(* IEC 61131-3 sources: 2026_Projet_YGO_ExcavatriceDragage/TOOLS/TEST_AUTO_CI/RESULTS/L_SIMULATION/tests (part 6) *)

(* ---- test_sim_operator_joystick.st ---- *)
(* T418 integration : vrais SimBench, FB_Joystick et homing, aucune logique machine remplacee.
   Temps explicite par scan : le DSL STruCpp interdit ADVANCE_TIME dans FOR. *)
SETUP
VAR
    bench : FB_SimBench;
    joy : FB_Joystick;
    home : FB_CycleMachineHoming;
    cfg : ST_fbJoystick_Cfg;
    diagOk : ST_Diag_Device;
    nx : INT := 5000;
    ny : INT := 5000;
    raw1 : UDINT;
    raw2 : UDINT;
    sourceSelected : BOOL;
    selectedX : INT;
    selectedY : INT;
    selectedButton : BOOL;
    previousButton : BOOL;
    buttonEdges : INT;
END_VAR
END_SETUP
TEST 'TC-T418-INT-001 Geste complet avec vrai joystick'
nx := 5000; ny := 5000; raw1 := 0; raw2 := 0; previousButton := FALSE; buttonEdges := 0;
bench.Enable := TRUE; joy.Enable := TRUE; joy.ArmingPermit := TRUE; diagOk.Operational := TRUE;
joy.BusCanOpenOP := diagOk; joy.JoystickOP := diagOk; home.Enable := TRUE; home.BootReady := TRUE;
home.Mode := E_Mode.MAINT_N1; home.BucketOffsetValid := TRUE; home.WinchesMechanicallyStopped := TRUE;
ADVANCE_TIME(10000000);
bench(RawPosM1 := raw1, RawPosM2 := raw2);
joy(RawX := bench.Operator.JoyXRaw_ANA1, RawY := bench.Operator.JoyYRaw_ANA2, RawButton := bench.Operator.JoyBtnRaw, Cfg := cfg, NeutralXMem := nx, NeutralYMem := ny);
home(DeadmanArmed := joy.DeadmanArmed, JoystickDeflected := NOT joy.AtNeutralXY, JoystickPull := joy.AxisCmdY.DirectionPositive, JoystickPush := joy.AxisCmdY.DirectionNegative, BtnValidation := bench.Operator.JoyBtnRaw);
IF bench.Operator.JoyBtnRaw AND NOT previousButton THEN buttonEdges := buttonEdges + 1; END_IF; previousButton := bench.Operator.JoyBtnRaw;
bench.SimJoystickRight_Fwd_MAINT_Active := TRUE;
ADVANCE_TIME(10000000);
bench(RawPosM1 := raw1, RawPosM2 := raw2);
joy(RawX := bench.Operator.JoyXRaw_ANA1, RawY := bench.Operator.JoyYRaw_ANA2, RawButton := bench.Operator.JoyBtnRaw, Cfg := cfg, NeutralXMem := nx, NeutralYMem := ny);
home(DeadmanArmed := joy.DeadmanArmed, JoystickDeflected := NOT joy.AtNeutralXY, JoystickPull := joy.AxisCmdY.DirectionPositive, JoystickPush := joy.AxisCmdY.DirectionNegative, BtnValidation := bench.Operator.JoyBtnRaw);
IF bench.Operator.JoyBtnRaw AND NOT previousButton THEN buttonEdges := buttonEdges + 1; END_IF; previousButton := bench.Operator.JoyBtnRaw;
ASSERT_EQ(bench.Operator.JoyXRaw_ANA1, 5000, 'Neutre pendant pre-appui');
ADVANCE_TIME(10000000);
bench(RawPosM1 := raw1, RawPosM2 := raw2);
joy(RawX := bench.Operator.JoyXRaw_ANA1, RawY := bench.Operator.JoyYRaw_ANA2, RawButton := bench.Operator.JoyBtnRaw, Cfg := cfg, NeutralXMem := nx, NeutralYMem := ny);
home(DeadmanArmed := joy.DeadmanArmed, JoystickDeflected := NOT joy.AtNeutralXY, JoystickPull := joy.AxisCmdY.DirectionPositive, JoystickPush := joy.AxisCmdY.DirectionNegative, BtnValidation := bench.Operator.JoyBtnRaw);
IF bench.Operator.JoyBtnRaw AND NOT previousButton THEN buttonEdges := buttonEdges + 1; END_IF; previousButton := bench.Operator.JoyBtnRaw;
ASSERT_EQ(bench.Operator.JoyXRaw_ANA1, 5000, 'Neutre pendant pre-appui');
ADVANCE_TIME(10000000);
bench(RawPosM1 := raw1, RawPosM2 := raw2);
joy(RawX := bench.Operator.JoyXRaw_ANA1, RawY := bench.Operator.JoyYRaw_ANA2, RawButton := bench.Operator.JoyBtnRaw, Cfg := cfg, NeutralXMem := nx, NeutralYMem := ny);
home(DeadmanArmed := joy.DeadmanArmed, JoystickDeflected := NOT joy.AtNeutralXY, JoystickPull := joy.AxisCmdY.DirectionPositive, JoystickPush := joy.AxisCmdY.DirectionNegative, BtnValidation := bench.Operator.JoyBtnRaw);
IF bench.Operator.JoyBtnRaw AND NOT previousButton THEN buttonEdges := buttonEdges + 1; END_IF; previousButton := bench.Operator.JoyBtnRaw;
ASSERT_EQ(bench.Operator.JoyXRaw_ANA1, 5000, 'Neutre pendant pre-appui');
ADVANCE_TIME(10000000);
bench(RawPosM1 := raw1, RawPosM2 := raw2);
joy(RawX := bench.Operator.JoyXRaw_ANA1, RawY := bench.Operator.JoyYRaw_ANA2, RawButton := bench.Operator.JoyBtnRaw, Cfg := cfg, NeutralXMem := nx, NeutralYMem := ny);
home(DeadmanArmed := joy.DeadmanArmed, JoystickDeflected := NOT joy.AtNeutralXY, JoystickPull := joy.AxisCmdY.DirectionPositive, JoystickPush := joy.AxisCmdY.DirectionNegative, BtnValidation := bench.Operator.JoyBtnRaw);
IF bench.Operator.JoyBtnRaw AND NOT previousButton THEN buttonEdges := buttonEdges + 1; END_IF; previousButton := bench.Operator.JoyBtnRaw;
ASSERT_EQ(bench.Operator.JoyXRaw_ANA1, 5000, 'Neutre pendant pre-appui');
ADVANCE_TIME(10000000);
bench(RawPosM1 := raw1, RawPosM2 := raw2);
joy(RawX := bench.Operator.JoyXRaw_ANA1, RawY := bench.Operator.JoyYRaw_ANA2, RawButton := bench.Operator.JoyBtnRaw, Cfg := cfg, NeutralXMem := nx, NeutralYMem := ny);
home(DeadmanArmed := joy.DeadmanArmed, JoystickDeflected := NOT joy.AtNeutralXY, JoystickPull := joy.AxisCmdY.DirectionPositive, JoystickPush := joy.AxisCmdY.DirectionNegative, BtnValidation := bench.Operator.JoyBtnRaw);
IF bench.Operator.JoyBtnRaw AND NOT previousButton THEN buttonEdges := buttonEdges + 1; END_IF; previousButton := bench.Operator.JoyBtnRaw;
ASSERT_EQ(bench.Operator.JoyXRaw_ANA1, 5000, 'Neutre pendant pre-appui');
ADVANCE_TIME(10000000);
bench(RawPosM1 := raw1, RawPosM2 := raw2);
joy(RawX := bench.Operator.JoyXRaw_ANA1, RawY := bench.Operator.JoyYRaw_ANA2, RawButton := bench.Operator.JoyBtnRaw, Cfg := cfg, NeutralXMem := nx, NeutralYMem := ny);
home(DeadmanArmed := joy.DeadmanArmed, JoystickDeflected := NOT joy.AtNeutralXY, JoystickPull := joy.AxisCmdY.DirectionPositive, JoystickPush := joy.AxisCmdY.DirectionNegative, BtnValidation := bench.Operator.JoyBtnRaw);
IF bench.Operator.JoyBtnRaw AND NOT previousButton THEN buttonEdges := buttonEdges + 1; END_IF; previousButton := bench.Operator.JoyBtnRaw;
ASSERT_EQ(bench.Operator.JoyXRaw_ANA1, 5000, 'Neutre pendant pre-appui');
ADVANCE_TIME(10000000);
bench(RawPosM1 := raw1, RawPosM2 := raw2);
joy(RawX := bench.Operator.JoyXRaw_ANA1, RawY := bench.Operator.JoyYRaw_ANA2, RawButton := bench.Operator.JoyBtnRaw, Cfg := cfg, NeutralXMem := nx, NeutralYMem := ny);
home(DeadmanArmed := joy.DeadmanArmed, JoystickDeflected := NOT joy.AtNeutralXY, JoystickPull := joy.AxisCmdY.DirectionPositive, JoystickPush := joy.AxisCmdY.DirectionNegative, BtnValidation := bench.Operator.JoyBtnRaw);
IF bench.Operator.JoyBtnRaw AND NOT previousButton THEN buttonEdges := buttonEdges + 1; END_IF; previousButton := bench.Operator.JoyBtnRaw;
ASSERT_EQ(bench.Operator.JoyXRaw_ANA1, 5000, 'Neutre pendant pre-appui');
ADVANCE_TIME(10000000);
bench(RawPosM1 := raw1, RawPosM2 := raw2);
joy(RawX := bench.Operator.JoyXRaw_ANA1, RawY := bench.Operator.JoyYRaw_ANA2, RawButton := bench.Operator.JoyBtnRaw, Cfg := cfg, NeutralXMem := nx, NeutralYMem := ny);
home(DeadmanArmed := joy.DeadmanArmed, JoystickDeflected := NOT joy.AtNeutralXY, JoystickPull := joy.AxisCmdY.DirectionPositive, JoystickPush := joy.AxisCmdY.DirectionNegative, BtnValidation := bench.Operator.JoyBtnRaw);
IF bench.Operator.JoyBtnRaw AND NOT previousButton THEN buttonEdges := buttonEdges + 1; END_IF; previousButton := bench.Operator.JoyBtnRaw;
ASSERT_EQ(bench.Operator.JoyXRaw_ANA1, 5000, 'Neutre pendant pre-appui');
ADVANCE_TIME(10000000);
bench(RawPosM1 := raw1, RawPosM2 := raw2);
joy(RawX := bench.Operator.JoyXRaw_ANA1, RawY := bench.Operator.JoyYRaw_ANA2, RawButton := bench.Operator.JoyBtnRaw, Cfg := cfg, NeutralXMem := nx, NeutralYMem := ny);
home(DeadmanArmed := joy.DeadmanArmed, JoystickDeflected := NOT joy.AtNeutralXY, JoystickPull := joy.AxisCmdY.DirectionPositive, JoystickPush := joy.AxisCmdY.DirectionNegative, BtnValidation := bench.Operator.JoyBtnRaw);
IF bench.Operator.JoyBtnRaw AND NOT previousButton THEN buttonEdges := buttonEdges + 1; END_IF; previousButton := bench.Operator.JoyBtnRaw;
ASSERT_EQ(bench.Operator.JoyXRaw_ANA1, 5000, 'Neutre pendant pre-appui');
ADVANCE_TIME(10000000);
bench(RawPosM1 := raw1, RawPosM2 := raw2);
joy(RawX := bench.Operator.JoyXRaw_ANA1, RawY := bench.Operator.JoyYRaw_ANA2, RawButton := bench.Operator.JoyBtnRaw, Cfg := cfg, NeutralXMem := nx, NeutralYMem := ny);
home(DeadmanArmed := joy.DeadmanArmed, JoystickDeflected := NOT joy.AtNeutralXY, JoystickPull := joy.AxisCmdY.DirectionPositive, JoystickPush := joy.AxisCmdY.DirectionNegative, BtnValidation := bench.Operator.JoyBtnRaw);
IF bench.Operator.JoyBtnRaw AND NOT previousButton THEN buttonEdges := buttonEdges + 1; END_IF; previousButton := bench.Operator.JoyBtnRaw;
ASSERT_EQ(bench.Operator.JoyXRaw_ANA1, 5000, 'Neutre pendant pre-appui');
ADVANCE_TIME(10000000);
bench(RawPosM1 := raw1, RawPosM2 := raw2);
joy(RawX := bench.Operator.JoyXRaw_ANA1, RawY := bench.Operator.JoyYRaw_ANA2, RawButton := bench.Operator.JoyBtnRaw, Cfg := cfg, NeutralXMem := nx, NeutralYMem := ny);
home(DeadmanArmed := joy.DeadmanArmed, JoystickDeflected := NOT joy.AtNeutralXY, JoystickPull := joy.AxisCmdY.DirectionPositive, JoystickPush := joy.AxisCmdY.DirectionNegative, BtnValidation := bench.Operator.JoyBtnRaw);
IF bench.Operator.JoyBtnRaw AND NOT previousButton THEN buttonEdges := buttonEdges + 1; END_IF; previousButton := bench.Operator.JoyBtnRaw;
ADVANCE_TIME(10000000);
bench(RawPosM1 := raw1, RawPosM2 := raw2);
joy(RawX := bench.Operator.JoyXRaw_ANA1, RawY := bench.Operator.JoyYRaw_ANA2, RawButton := bench.Operator.JoyBtnRaw, Cfg := cfg, NeutralXMem := nx, NeutralYMem := ny);
home(DeadmanArmed := joy.DeadmanArmed, JoystickDeflected := NOT joy.AtNeutralXY, JoystickPull := joy.AxisCmdY.DirectionPositive, JoystickPush := joy.AxisCmdY.DirectionNegative, BtnValidation := bench.Operator.JoyBtnRaw);
IF bench.Operator.JoyBtnRaw AND NOT previousButton THEN buttonEdges := buttonEdges + 1; END_IF; previousButton := bench.Operator.JoyBtnRaw;
ADVANCE_TIME(10000000);
bench(RawPosM1 := raw1, RawPosM2 := raw2);
joy(RawX := bench.Operator.JoyXRaw_ANA1, RawY := bench.Operator.JoyYRaw_ANA2, RawButton := bench.Operator.JoyBtnRaw, Cfg := cfg, NeutralXMem := nx, NeutralYMem := ny);
home(DeadmanArmed := joy.DeadmanArmed, JoystickDeflected := NOT joy.AtNeutralXY, JoystickPull := joy.AxisCmdY.DirectionPositive, JoystickPush := joy.AxisCmdY.DirectionNegative, BtnValidation := bench.Operator.JoyBtnRaw);
IF bench.Operator.JoyBtnRaw AND NOT previousButton THEN buttonEdges := buttonEdges + 1; END_IF; previousButton := bench.Operator.JoyBtnRaw;
ADVANCE_TIME(10000000);
bench(RawPosM1 := raw1, RawPosM2 := raw2);
joy(RawX := bench.Operator.JoyXRaw_ANA1, RawY := bench.Operator.JoyYRaw_ANA2, RawButton := bench.Operator.JoyBtnRaw, Cfg := cfg, NeutralXMem := nx, NeutralYMem := ny);
home(DeadmanArmed := joy.DeadmanArmed, JoystickDeflected := NOT joy.AtNeutralXY, JoystickPull := joy.AxisCmdY.DirectionPositive, JoystickPush := joy.AxisCmdY.DirectionNegative, BtnValidation := bench.Operator.JoyBtnRaw);
IF bench.Operator.JoyBtnRaw AND NOT previousButton THEN buttonEdges := buttonEdges + 1; END_IF; previousButton := bench.Operator.JoyBtnRaw;
ASSERT_TRUE(joy.DeadmanArmed, 'Le vrai joystick arme par maintien');
ADVANCE_TIME(10000000);
bench(RawPosM1 := raw1, RawPosM2 := raw2);
joy(RawX := bench.Operator.JoyXRaw_ANA1, RawY := bench.Operator.JoyYRaw_ANA2, RawButton := bench.Operator.JoyBtnRaw, Cfg := cfg, NeutralXMem := nx, NeutralYMem := ny);
home(DeadmanArmed := joy.DeadmanArmed, JoystickDeflected := NOT joy.AtNeutralXY, JoystickPull := joy.AxisCmdY.DirectionPositive, JoystickPush := joy.AxisCmdY.DirectionNegative, BtnValidation := bench.Operator.JoyBtnRaw);
IF bench.Operator.JoyBtnRaw AND NOT previousButton THEN buttonEdges := buttonEdges + 1; END_IF; previousButton := bench.Operator.JoyBtnRaw;
ADVANCE_TIME(10000000);
bench(RawPosM1 := raw1, RawPosM2 := raw2);
joy(RawX := bench.Operator.JoyXRaw_ANA1, RawY := bench.Operator.JoyYRaw_ANA2, RawButton := bench.Operator.JoyBtnRaw, Cfg := cfg, NeutralXMem := nx, NeutralYMem := ny);
home(DeadmanArmed := joy.DeadmanArmed, JoystickDeflected := NOT joy.AtNeutralXY, JoystickPull := joy.AxisCmdY.DirectionPositive, JoystickPush := joy.AxisCmdY.DirectionNegative, BtnValidation := bench.Operator.JoyBtnRaw);
IF bench.Operator.JoyBtnRaw AND NOT previousButton THEN buttonEdges := buttonEdges + 1; END_IF; previousButton := bench.Operator.JoyBtnRaw;
ADVANCE_TIME(10000000);
bench(RawPosM1 := raw1, RawPosM2 := raw2);
joy(RawX := bench.Operator.JoyXRaw_ANA1, RawY := bench.Operator.JoyYRaw_ANA2, RawButton := bench.Operator.JoyBtnRaw, Cfg := cfg, NeutralXMem := nx, NeutralYMem := ny);
home(DeadmanArmed := joy.DeadmanArmed, JoystickDeflected := NOT joy.AtNeutralXY, JoystickPull := joy.AxisCmdY.DirectionPositive, JoystickPush := joy.AxisCmdY.DirectionNegative, BtnValidation := bench.Operator.JoyBtnRaw);
IF bench.Operator.JoyBtnRaw AND NOT previousButton THEN buttonEdges := buttonEdges + 1; END_IF; previousButton := bench.Operator.JoyBtnRaw;
ADVANCE_TIME(10000000);
bench(RawPosM1 := raw1, RawPosM2 := raw2);
joy(RawX := bench.Operator.JoyXRaw_ANA1, RawY := bench.Operator.JoyYRaw_ANA2, RawButton := bench.Operator.JoyBtnRaw, Cfg := cfg, NeutralXMem := nx, NeutralYMem := ny);
home(DeadmanArmed := joy.DeadmanArmed, JoystickDeflected := NOT joy.AtNeutralXY, JoystickPull := joy.AxisCmdY.DirectionPositive, JoystickPush := joy.AxisCmdY.DirectionNegative, BtnValidation := bench.Operator.JoyBtnRaw);
IF bench.Operator.JoyBtnRaw AND NOT previousButton THEN buttonEdges := buttonEdges + 1; END_IF; previousButton := bench.Operator.JoyBtnRaw;
ADVANCE_TIME(10000000);
bench(RawPosM1 := raw1, RawPosM2 := raw2);
joy(RawX := bench.Operator.JoyXRaw_ANA1, RawY := bench.Operator.JoyYRaw_ANA2, RawButton := bench.Operator.JoyBtnRaw, Cfg := cfg, NeutralXMem := nx, NeutralYMem := ny);
home(DeadmanArmed := joy.DeadmanArmed, JoystickDeflected := NOT joy.AtNeutralXY, JoystickPull := joy.AxisCmdY.DirectionPositive, JoystickPush := joy.AxisCmdY.DirectionNegative, BtnValidation := bench.Operator.JoyBtnRaw);
IF bench.Operator.JoyBtnRaw AND NOT previousButton THEN buttonEdges := buttonEdges + 1; END_IF; previousButton := bench.Operator.JoyBtnRaw;
ADVANCE_TIME(10000000);
bench(RawPosM1 := raw1, RawPosM2 := raw2);
joy(RawX := bench.Operator.JoyXRaw_ANA1, RawY := bench.Operator.JoyYRaw_ANA2, RawButton := bench.Operator.JoyBtnRaw, Cfg := cfg, NeutralXMem := nx, NeutralYMem := ny);
home(DeadmanArmed := joy.DeadmanArmed, JoystickDeflected := NOT joy.AtNeutralXY, JoystickPull := joy.AxisCmdY.DirectionPositive, JoystickPush := joy.AxisCmdY.DirectionNegative, BtnValidation := bench.Operator.JoyBtnRaw);
IF bench.Operator.JoyBtnRaw AND NOT previousButton THEN buttonEdges := buttonEdges + 1; END_IF; previousButton := bench.Operator.JoyBtnRaw;
ADVANCE_TIME(10000000);
bench(RawPosM1 := raw1, RawPosM2 := raw2);
joy(RawX := bench.Operator.JoyXRaw_ANA1, RawY := bench.Operator.JoyYRaw_ANA2, RawButton := bench.Operator.JoyBtnRaw, Cfg := cfg, NeutralXMem := nx, NeutralYMem := ny);
home(DeadmanArmed := joy.DeadmanArmed, JoystickDeflected := NOT joy.AtNeutralXY, JoystickPull := joy.AxisCmdY.DirectionPositive, JoystickPush := joy.AxisCmdY.DirectionNegative, BtnValidation := bench.Operator.JoyBtnRaw);
IF bench.Operator.JoyBtnRaw AND NOT previousButton THEN buttonEdges := buttonEdges + 1; END_IF; previousButton := bench.Operator.JoyBtnRaw;
ADVANCE_TIME(10000000);
bench(RawPosM1 := raw1, RawPosM2 := raw2);
joy(RawX := bench.Operator.JoyXRaw_ANA1, RawY := bench.Operator.JoyYRaw_ANA2, RawButton := bench.Operator.JoyBtnRaw, Cfg := cfg, NeutralXMem := nx, NeutralYMem := ny);
home(DeadmanArmed := joy.DeadmanArmed, JoystickDeflected := NOT joy.AtNeutralXY, JoystickPull := joy.AxisCmdY.DirectionPositive, JoystickPush := joy.AxisCmdY.DirectionNegative, BtnValidation := bench.Operator.JoyBtnRaw);
IF bench.Operator.JoyBtnRaw AND NOT previousButton THEN buttonEdges := buttonEdges + 1; END_IF; previousButton := bench.Operator.JoyBtnRaw;
ADVANCE_TIME(10000000);
bench(RawPosM1 := raw1, RawPosM2 := raw2);
joy(RawX := bench.Operator.JoyXRaw_ANA1, RawY := bench.Operator.JoyYRaw_ANA2, RawButton := bench.Operator.JoyBtnRaw, Cfg := cfg, NeutralXMem := nx, NeutralYMem := ny);
home(DeadmanArmed := joy.DeadmanArmed, JoystickDeflected := NOT joy.AtNeutralXY, JoystickPull := joy.AxisCmdY.DirectionPositive, JoystickPush := joy.AxisCmdY.DirectionNegative, BtnValidation := bench.Operator.JoyBtnRaw);
IF bench.Operator.JoyBtnRaw AND NOT previousButton THEN buttonEdges := buttonEdges + 1; END_IF; previousButton := bench.Operator.JoyBtnRaw;
ADVANCE_TIME(10000000);
bench(RawPosM1 := raw1, RawPosM2 := raw2);
joy(RawX := bench.Operator.JoyXRaw_ANA1, RawY := bench.Operator.JoyYRaw_ANA2, RawButton := bench.Operator.JoyBtnRaw, Cfg := cfg, NeutralXMem := nx, NeutralYMem := ny);
home(DeadmanArmed := joy.DeadmanArmed, JoystickDeflected := NOT joy.AtNeutralXY, JoystickPull := joy.AxisCmdY.DirectionPositive, JoystickPush := joy.AxisCmdY.DirectionNegative, BtnValidation := bench.Operator.JoyBtnRaw);
IF bench.Operator.JoyBtnRaw AND NOT previousButton THEN buttonEdges := buttonEdges + 1; END_IF; previousButton := bench.Operator.JoyBtnRaw;
ADVANCE_TIME(10000000);
bench(RawPosM1 := raw1, RawPosM2 := raw2);
joy(RawX := bench.Operator.JoyXRaw_ANA1, RawY := bench.Operator.JoyYRaw_ANA2, RawButton := bench.Operator.JoyBtnRaw, Cfg := cfg, NeutralXMem := nx, NeutralYMem := ny);
home(DeadmanArmed := joy.DeadmanArmed, JoystickDeflected := NOT joy.AtNeutralXY, JoystickPull := joy.AxisCmdY.DirectionPositive, JoystickPush := joy.AxisCmdY.DirectionNegative, BtnValidation := bench.Operator.JoyBtnRaw);
IF bench.Operator.JoyBtnRaw AND NOT previousButton THEN buttonEdges := buttonEdges + 1; END_IF; previousButton := bench.Operator.JoyBtnRaw;
ADVANCE_TIME(10000000);
bench(RawPosM1 := raw1, RawPosM2 := raw2);
joy(RawX := bench.Operator.JoyXRaw_ANA1, RawY := bench.Operator.JoyYRaw_ANA2, RawButton := bench.Operator.JoyBtnRaw, Cfg := cfg, NeutralXMem := nx, NeutralYMem := ny);
home(DeadmanArmed := joy.DeadmanArmed, JoystickDeflected := NOT joy.AtNeutralXY, JoystickPull := joy.AxisCmdY.DirectionPositive, JoystickPush := joy.AxisCmdY.DirectionNegative, BtnValidation := bench.Operator.JoyBtnRaw);
IF bench.Operator.JoyBtnRaw AND NOT previousButton THEN buttonEdges := buttonEdges + 1; END_IF; previousButton := bench.Operator.JoyBtnRaw;
ADVANCE_TIME(10000000);
bench(RawPosM1 := raw1, RawPosM2 := raw2);
joy(RawX := bench.Operator.JoyXRaw_ANA1, RawY := bench.Operator.JoyYRaw_ANA2, RawButton := bench.Operator.JoyBtnRaw, Cfg := cfg, NeutralXMem := nx, NeutralYMem := ny);
home(DeadmanArmed := joy.DeadmanArmed, JoystickDeflected := NOT joy.AtNeutralXY, JoystickPull := joy.AxisCmdY.DirectionPositive, JoystickPush := joy.AxisCmdY.DirectionNegative, BtnValidation := bench.Operator.JoyBtnRaw);
IF bench.Operator.JoyBtnRaw AND NOT previousButton THEN buttonEdges := buttonEdges + 1; END_IF; previousButton := bench.Operator.JoyBtnRaw;
ADVANCE_TIME(10000000);
bench(RawPosM1 := raw1, RawPosM2 := raw2);
joy(RawX := bench.Operator.JoyXRaw_ANA1, RawY := bench.Operator.JoyYRaw_ANA2, RawButton := bench.Operator.JoyBtnRaw, Cfg := cfg, NeutralXMem := nx, NeutralYMem := ny);
home(DeadmanArmed := joy.DeadmanArmed, JoystickDeflected := NOT joy.AtNeutralXY, JoystickPull := joy.AxisCmdY.DirectionPositive, JoystickPush := joy.AxisCmdY.DirectionNegative, BtnValidation := bench.Operator.JoyBtnRaw);
IF bench.Operator.JoyBtnRaw AND NOT previousButton THEN buttonEdges := buttonEdges + 1; END_IF; previousButton := bench.Operator.JoyBtnRaw;
ADVANCE_TIME(10000000);
bench(RawPosM1 := raw1, RawPosM2 := raw2);
joy(RawX := bench.Operator.JoyXRaw_ANA1, RawY := bench.Operator.JoyYRaw_ANA2, RawButton := bench.Operator.JoyBtnRaw, Cfg := cfg, NeutralXMem := nx, NeutralYMem := ny);
home(DeadmanArmed := joy.DeadmanArmed, JoystickDeflected := NOT joy.AtNeutralXY, JoystickPull := joy.AxisCmdY.DirectionPositive, JoystickPush := joy.AxisCmdY.DirectionNegative, BtnValidation := bench.Operator.JoyBtnRaw);
IF bench.Operator.JoyBtnRaw AND NOT previousButton THEN buttonEdges := buttonEdges + 1; END_IF; previousButton := bench.Operator.JoyBtnRaw;
ADVANCE_TIME(10000000);
bench(RawPosM1 := raw1, RawPosM2 := raw2);
joy(RawX := bench.Operator.JoyXRaw_ANA1, RawY := bench.Operator.JoyYRaw_ANA2, RawButton := bench.Operator.JoyBtnRaw, Cfg := cfg, NeutralXMem := nx, NeutralYMem := ny);
home(DeadmanArmed := joy.DeadmanArmed, JoystickDeflected := NOT joy.AtNeutralXY, JoystickPull := joy.AxisCmdY.DirectionPositive, JoystickPush := joy.AxisCmdY.DirectionNegative, BtnValidation := bench.Operator.JoyBtnRaw);
IF bench.Operator.JoyBtnRaw AND NOT previousButton THEN buttonEdges := buttonEdges + 1; END_IF; previousButton := bench.Operator.JoyBtnRaw;
ADVANCE_TIME(10000000);
bench(RawPosM1 := raw1, RawPosM2 := raw2);
joy(RawX := bench.Operator.JoyXRaw_ANA1, RawY := bench.Operator.JoyYRaw_ANA2, RawButton := bench.Operator.JoyBtnRaw, Cfg := cfg, NeutralXMem := nx, NeutralYMem := ny);
home(DeadmanArmed := joy.DeadmanArmed, JoystickDeflected := NOT joy.AtNeutralXY, JoystickPull := joy.AxisCmdY.DirectionPositive, JoystickPush := joy.AxisCmdY.DirectionNegative, BtnValidation := bench.Operator.JoyBtnRaw);
IF bench.Operator.JoyBtnRaw AND NOT previousButton THEN buttonEdges := buttonEdges + 1; END_IF; previousButton := bench.Operator.JoyBtnRaw;
ADVANCE_TIME(10000000);
bench(RawPosM1 := raw1, RawPosM2 := raw2);
joy(RawX := bench.Operator.JoyXRaw_ANA1, RawY := bench.Operator.JoyYRaw_ANA2, RawButton := bench.Operator.JoyBtnRaw, Cfg := cfg, NeutralXMem := nx, NeutralYMem := ny);
home(DeadmanArmed := joy.DeadmanArmed, JoystickDeflected := NOT joy.AtNeutralXY, JoystickPull := joy.AxisCmdY.DirectionPositive, JoystickPush := joy.AxisCmdY.DirectionNegative, BtnValidation := bench.Operator.JoyBtnRaw);
IF bench.Operator.JoyBtnRaw AND NOT previousButton THEN buttonEdges := buttonEdges + 1; END_IF; previousButton := bench.Operator.JoyBtnRaw;
ADVANCE_TIME(10000000);
bench(RawPosM1 := raw1, RawPosM2 := raw2);
joy(RawX := bench.Operator.JoyXRaw_ANA1, RawY := bench.Operator.JoyYRaw_ANA2, RawButton := bench.Operator.JoyBtnRaw, Cfg := cfg, NeutralXMem := nx, NeutralYMem := ny);
home(DeadmanArmed := joy.DeadmanArmed, JoystickDeflected := NOT joy.AtNeutralXY, JoystickPull := joy.AxisCmdY.DirectionPositive, JoystickPush := joy.AxisCmdY.DirectionNegative, BtnValidation := bench.Operator.JoyBtnRaw);
IF bench.Operator.JoyBtnRaw AND NOT previousButton THEN buttonEdges := buttonEdges + 1; END_IF; previousButton := bench.Operator.JoyBtnRaw;
ADVANCE_TIME(10000000);
bench(RawPosM1 := raw1, RawPosM2 := raw2);
joy(RawX := bench.Operator.JoyXRaw_ANA1, RawY := bench.Operator.JoyYRaw_ANA2, RawButton := bench.Operator.JoyBtnRaw, Cfg := cfg, NeutralXMem := nx, NeutralYMem := ny);
home(DeadmanArmed := joy.DeadmanArmed, JoystickDeflected := NOT joy.AtNeutralXY, JoystickPull := joy.AxisCmdY.DirectionPositive, JoystickPush := joy.AxisCmdY.DirectionNegative, BtnValidation := bench.Operator.JoyBtnRaw);
IF bench.Operator.JoyBtnRaw AND NOT previousButton THEN buttonEdges := buttonEdges + 1; END_IF; previousButton := bench.Operator.JoyBtnRaw;
ADVANCE_TIME(10000000);
bench(RawPosM1 := raw1, RawPosM2 := raw2);
joy(RawX := bench.Operator.JoyXRaw_ANA1, RawY := bench.Operator.JoyYRaw_ANA2, RawButton := bench.Operator.JoyBtnRaw, Cfg := cfg, NeutralXMem := nx, NeutralYMem := ny);
home(DeadmanArmed := joy.DeadmanArmed, JoystickDeflected := NOT joy.AtNeutralXY, JoystickPull := joy.AxisCmdY.DirectionPositive, JoystickPush := joy.AxisCmdY.DirectionNegative, BtnValidation := bench.Operator.JoyBtnRaw);
IF bench.Operator.JoyBtnRaw AND NOT previousButton THEN buttonEdges := buttonEdges + 1; END_IF; previousButton := bench.Operator.JoyBtnRaw;
ADVANCE_TIME(10000000);
bench(RawPosM1 := raw1, RawPosM2 := raw2);
joy(RawX := bench.Operator.JoyXRaw_ANA1, RawY := bench.Operator.JoyYRaw_ANA2, RawButton := bench.Operator.JoyBtnRaw, Cfg := cfg, NeutralXMem := nx, NeutralYMem := ny);
home(DeadmanArmed := joy.DeadmanArmed, JoystickDeflected := NOT joy.AtNeutralXY, JoystickPull := joy.AxisCmdY.DirectionPositive, JoystickPush := joy.AxisCmdY.DirectionNegative, BtnValidation := bench.Operator.JoyBtnRaw);
IF bench.Operator.JoyBtnRaw AND NOT previousButton THEN buttonEdges := buttonEdges + 1; END_IF; previousButton := bench.Operator.JoyBtnRaw;
ADVANCE_TIME(10000000);
bench(RawPosM1 := raw1, RawPosM2 := raw2);
joy(RawX := bench.Operator.JoyXRaw_ANA1, RawY := bench.Operator.JoyYRaw_ANA2, RawButton := bench.Operator.JoyBtnRaw, Cfg := cfg, NeutralXMem := nx, NeutralYMem := ny);
home(DeadmanArmed := joy.DeadmanArmed, JoystickDeflected := NOT joy.AtNeutralXY, JoystickPull := joy.AxisCmdY.DirectionPositive, JoystickPush := joy.AxisCmdY.DirectionNegative, BtnValidation := bench.Operator.JoyBtnRaw);
IF bench.Operator.JoyBtnRaw AND NOT previousButton THEN buttonEdges := buttonEdges + 1; END_IF; previousButton := bench.Operator.JoyBtnRaw;
ADVANCE_TIME(10000000);
bench(RawPosM1 := raw1, RawPosM2 := raw2);
joy(RawX := bench.Operator.JoyXRaw_ANA1, RawY := bench.Operator.JoyYRaw_ANA2, RawButton := bench.Operator.JoyBtnRaw, Cfg := cfg, NeutralXMem := nx, NeutralYMem := ny);
home(DeadmanArmed := joy.DeadmanArmed, JoystickDeflected := NOT joy.AtNeutralXY, JoystickPull := joy.AxisCmdY.DirectionPositive, JoystickPush := joy.AxisCmdY.DirectionNegative, BtnValidation := bench.Operator.JoyBtnRaw);
IF bench.Operator.JoyBtnRaw AND NOT previousButton THEN buttonEdges := buttonEdges + 1; END_IF; previousButton := bench.Operator.JoyBtnRaw;
ADVANCE_TIME(10000000);
bench(RawPosM1 := raw1, RawPosM2 := raw2);
joy(RawX := bench.Operator.JoyXRaw_ANA1, RawY := bench.Operator.JoyYRaw_ANA2, RawButton := bench.Operator.JoyBtnRaw, Cfg := cfg, NeutralXMem := nx, NeutralYMem := ny);
home(DeadmanArmed := joy.DeadmanArmed, JoystickDeflected := NOT joy.AtNeutralXY, JoystickPull := joy.AxisCmdY.DirectionPositive, JoystickPush := joy.AxisCmdY.DirectionNegative, BtnValidation := bench.Operator.JoyBtnRaw);
IF bench.Operator.JoyBtnRaw AND NOT previousButton THEN buttonEdges := buttonEdges + 1; END_IF; previousButton := bench.Operator.JoyBtnRaw;
ADVANCE_TIME(10000000);
bench(RawPosM1 := raw1, RawPosM2 := raw2);
joy(RawX := bench.Operator.JoyXRaw_ANA1, RawY := bench.Operator.JoyYRaw_ANA2, RawButton := bench.Operator.JoyBtnRaw, Cfg := cfg, NeutralXMem := nx, NeutralYMem := ny);
home(DeadmanArmed := joy.DeadmanArmed, JoystickDeflected := NOT joy.AtNeutralXY, JoystickPull := joy.AxisCmdY.DirectionPositive, JoystickPush := joy.AxisCmdY.DirectionNegative, BtnValidation := bench.Operator.JoyBtnRaw);
IF bench.Operator.JoyBtnRaw AND NOT previousButton THEN buttonEdges := buttonEdges + 1; END_IF; previousButton := bench.Operator.JoyBtnRaw;
ADVANCE_TIME(10000000);
bench(RawPosM1 := raw1, RawPosM2 := raw2);
joy(RawX := bench.Operator.JoyXRaw_ANA1, RawY := bench.Operator.JoyYRaw_ANA2, RawButton := bench.Operator.JoyBtnRaw, Cfg := cfg, NeutralXMem := nx, NeutralYMem := ny);
home(DeadmanArmed := joy.DeadmanArmed, JoystickDeflected := NOT joy.AtNeutralXY, JoystickPull := joy.AxisCmdY.DirectionPositive, JoystickPush := joy.AxisCmdY.DirectionNegative, BtnValidation := bench.Operator.JoyBtnRaw);
IF bench.Operator.JoyBtnRaw AND NOT previousButton THEN buttonEdges := buttonEdges + 1; END_IF; previousButton := bench.Operator.JoyBtnRaw;
ADVANCE_TIME(10000000);
bench(RawPosM1 := raw1, RawPosM2 := raw2);
joy(RawX := bench.Operator.JoyXRaw_ANA1, RawY := bench.Operator.JoyYRaw_ANA2, RawButton := bench.Operator.JoyBtnRaw, Cfg := cfg, NeutralXMem := nx, NeutralYMem := ny);
home(DeadmanArmed := joy.DeadmanArmed, JoystickDeflected := NOT joy.AtNeutralXY, JoystickPull := joy.AxisCmdY.DirectionPositive, JoystickPush := joy.AxisCmdY.DirectionNegative, BtnValidation := bench.Operator.JoyBtnRaw);
IF bench.Operator.JoyBtnRaw AND NOT previousButton THEN buttonEdges := buttonEdges + 1; END_IF; previousButton := bench.Operator.JoyBtnRaw;
ADVANCE_TIME(10000000);
bench(RawPosM1 := raw1, RawPosM2 := raw2);
joy(RawX := bench.Operator.JoyXRaw_ANA1, RawY := bench.Operator.JoyYRaw_ANA2, RawButton := bench.Operator.JoyBtnRaw, Cfg := cfg, NeutralXMem := nx, NeutralYMem := ny);
home(DeadmanArmed := joy.DeadmanArmed, JoystickDeflected := NOT joy.AtNeutralXY, JoystickPull := joy.AxisCmdY.DirectionPositive, JoystickPush := joy.AxisCmdY.DirectionNegative, BtnValidation := bench.Operator.JoyBtnRaw);
IF bench.Operator.JoyBtnRaw AND NOT previousButton THEN buttonEdges := buttonEdges + 1; END_IF; previousButton := bench.Operator.JoyBtnRaw;
ADVANCE_TIME(10000000);
bench(RawPosM1 := raw1, RawPosM2 := raw2);
joy(RawX := bench.Operator.JoyXRaw_ANA1, RawY := bench.Operator.JoyYRaw_ANA2, RawButton := bench.Operator.JoyBtnRaw, Cfg := cfg, NeutralXMem := nx, NeutralYMem := ny);
home(DeadmanArmed := joy.DeadmanArmed, JoystickDeflected := NOT joy.AtNeutralXY, JoystickPull := joy.AxisCmdY.DirectionPositive, JoystickPush := joy.AxisCmdY.DirectionNegative, BtnValidation := bench.Operator.JoyBtnRaw);
IF bench.Operator.JoyBtnRaw AND NOT previousButton THEN buttonEdges := buttonEdges + 1; END_IF; previousButton := bench.Operator.JoyBtnRaw;
ADVANCE_TIME(10000000);
bench(RawPosM1 := raw1, RawPosM2 := raw2);
joy(RawX := bench.Operator.JoyXRaw_ANA1, RawY := bench.Operator.JoyYRaw_ANA2, RawButton := bench.Operator.JoyBtnRaw, Cfg := cfg, NeutralXMem := nx, NeutralYMem := ny);
home(DeadmanArmed := joy.DeadmanArmed, JoystickDeflected := NOT joy.AtNeutralXY, JoystickPull := joy.AxisCmdY.DirectionPositive, JoystickPush := joy.AxisCmdY.DirectionNegative, BtnValidation := bench.Operator.JoyBtnRaw);
IF bench.Operator.JoyBtnRaw AND NOT previousButton THEN buttonEdges := buttonEdges + 1; END_IF; previousButton := bench.Operator.JoyBtnRaw;
ADVANCE_TIME(10000000);
bench(RawPosM1 := raw1, RawPosM2 := raw2);
joy(RawX := bench.Operator.JoyXRaw_ANA1, RawY := bench.Operator.JoyYRaw_ANA2, RawButton := bench.Operator.JoyBtnRaw, Cfg := cfg, NeutralXMem := nx, NeutralYMem := ny);
home(DeadmanArmed := joy.DeadmanArmed, JoystickDeflected := NOT joy.AtNeutralXY, JoystickPull := joy.AxisCmdY.DirectionPositive, JoystickPush := joy.AxisCmdY.DirectionNegative, BtnValidation := bench.Operator.JoyBtnRaw);
IF bench.Operator.JoyBtnRaw AND NOT previousButton THEN buttonEdges := buttonEdges + 1; END_IF; previousButton := bench.Operator.JoyBtnRaw;
ADVANCE_TIME(10000000);
bench(RawPosM1 := raw1, RawPosM2 := raw2);
joy(RawX := bench.Operator.JoyXRaw_ANA1, RawY := bench.Operator.JoyYRaw_ANA2, RawButton := bench.Operator.JoyBtnRaw, Cfg := cfg, NeutralXMem := nx, NeutralYMem := ny);
home(DeadmanArmed := joy.DeadmanArmed, JoystickDeflected := NOT joy.AtNeutralXY, JoystickPull := joy.AxisCmdY.DirectionPositive, JoystickPush := joy.AxisCmdY.DirectionNegative, BtnValidation := bench.Operator.JoyBtnRaw);
IF bench.Operator.JoyBtnRaw AND NOT previousButton THEN buttonEdges := buttonEdges + 1; END_IF; previousButton := bench.Operator.JoyBtnRaw;
ADVANCE_TIME(10000000);
bench(RawPosM1 := raw1, RawPosM2 := raw2);
joy(RawX := bench.Operator.JoyXRaw_ANA1, RawY := bench.Operator.JoyYRaw_ANA2, RawButton := bench.Operator.JoyBtnRaw, Cfg := cfg, NeutralXMem := nx, NeutralYMem := ny);
home(DeadmanArmed := joy.DeadmanArmed, JoystickDeflected := NOT joy.AtNeutralXY, JoystickPull := joy.AxisCmdY.DirectionPositive, JoystickPush := joy.AxisCmdY.DirectionNegative, BtnValidation := bench.Operator.JoyBtnRaw);
IF bench.Operator.JoyBtnRaw AND NOT previousButton THEN buttonEdges := buttonEdges + 1; END_IF; previousButton := bench.Operator.JoyBtnRaw;
ADVANCE_TIME(10000000);
bench(RawPosM1 := raw1, RawPosM2 := raw2);
joy(RawX := bench.Operator.JoyXRaw_ANA1, RawY := bench.Operator.JoyYRaw_ANA2, RawButton := bench.Operator.JoyBtnRaw, Cfg := cfg, NeutralXMem := nx, NeutralYMem := ny);
home(DeadmanArmed := joy.DeadmanArmed, JoystickDeflected := NOT joy.AtNeutralXY, JoystickPull := joy.AxisCmdY.DirectionPositive, JoystickPush := joy.AxisCmdY.DirectionNegative, BtnValidation := bench.Operator.JoyBtnRaw);
IF bench.Operator.JoyBtnRaw AND NOT previousButton THEN buttonEdges := buttonEdges + 1; END_IF; previousButton := bench.Operator.JoyBtnRaw;
ADVANCE_TIME(10000000);
bench(RawPosM1 := raw1, RawPosM2 := raw2);
joy(RawX := bench.Operator.JoyXRaw_ANA1, RawY := bench.Operator.JoyYRaw_ANA2, RawButton := bench.Operator.JoyBtnRaw, Cfg := cfg, NeutralXMem := nx, NeutralYMem := ny);
home(DeadmanArmed := joy.DeadmanArmed, JoystickDeflected := NOT joy.AtNeutralXY, JoystickPull := joy.AxisCmdY.DirectionPositive, JoystickPush := joy.AxisCmdY.DirectionNegative, BtnValidation := bench.Operator.JoyBtnRaw);
IF bench.Operator.JoyBtnRaw AND NOT previousButton THEN buttonEdges := buttonEdges + 1; END_IF; previousButton := bench.Operator.JoyBtnRaw;
ADVANCE_TIME(10000000);
bench(RawPosM1 := raw1, RawPosM2 := raw2);
joy(RawX := bench.Operator.JoyXRaw_ANA1, RawY := bench.Operator.JoyYRaw_ANA2, RawButton := bench.Operator.JoyBtnRaw, Cfg := cfg, NeutralXMem := nx, NeutralYMem := ny);
home(DeadmanArmed := joy.DeadmanArmed, JoystickDeflected := NOT joy.AtNeutralXY, JoystickPull := joy.AxisCmdY.DirectionPositive, JoystickPush := joy.AxisCmdY.DirectionNegative, BtnValidation := bench.Operator.JoyBtnRaw);
IF bench.Operator.JoyBtnRaw AND NOT previousButton THEN buttonEdges := buttonEdges + 1; END_IF; previousButton := bench.Operator.JoyBtnRaw;
ADVANCE_TIME(10000000);
bench(RawPosM1 := raw1, RawPosM2 := raw2);
joy(RawX := bench.Operator.JoyXRaw_ANA1, RawY := bench.Operator.JoyYRaw_ANA2, RawButton := bench.Operator.JoyBtnRaw, Cfg := cfg, NeutralXMem := nx, NeutralYMem := ny);
home(DeadmanArmed := joy.DeadmanArmed, JoystickDeflected := NOT joy.AtNeutralXY, JoystickPull := joy.AxisCmdY.DirectionPositive, JoystickPush := joy.AxisCmdY.DirectionNegative, BtnValidation := bench.Operator.JoyBtnRaw);
IF bench.Operator.JoyBtnRaw AND NOT previousButton THEN buttonEdges := buttonEdges + 1; END_IF; previousButton := bench.Operator.JoyBtnRaw;
ADVANCE_TIME(10000000);
bench(RawPosM1 := raw1, RawPosM2 := raw2);
joy(RawX := bench.Operator.JoyXRaw_ANA1, RawY := bench.Operator.JoyYRaw_ANA2, RawButton := bench.Operator.JoyBtnRaw, Cfg := cfg, NeutralXMem := nx, NeutralYMem := ny);
home(DeadmanArmed := joy.DeadmanArmed, JoystickDeflected := NOT joy.AtNeutralXY, JoystickPull := joy.AxisCmdY.DirectionPositive, JoystickPush := joy.AxisCmdY.DirectionNegative, BtnValidation := bench.Operator.JoyBtnRaw);
IF bench.Operator.JoyBtnRaw AND NOT previousButton THEN buttonEdges := buttonEdges + 1; END_IF; previousButton := bench.Operator.JoyBtnRaw;
ADVANCE_TIME(10000000);
bench(RawPosM1 := raw1, RawPosM2 := raw2);
joy(RawX := bench.Operator.JoyXRaw_ANA1, RawY := bench.Operator.JoyYRaw_ANA2, RawButton := bench.Operator.JoyBtnRaw, Cfg := cfg, NeutralXMem := nx, NeutralYMem := ny);
home(DeadmanArmed := joy.DeadmanArmed, JoystickDeflected := NOT joy.AtNeutralXY, JoystickPull := joy.AxisCmdY.DirectionPositive, JoystickPush := joy.AxisCmdY.DirectionNegative, BtnValidation := bench.Operator.JoyBtnRaw);
IF bench.Operator.JoyBtnRaw AND NOT previousButton THEN buttonEdges := buttonEdges + 1; END_IF; previousButton := bench.Operator.JoyBtnRaw;
ADVANCE_TIME(10000000);
bench(RawPosM1 := raw1, RawPosM2 := raw2);
joy(RawX := bench.Operator.JoyXRaw_ANA1, RawY := bench.Operator.JoyYRaw_ANA2, RawButton := bench.Operator.JoyBtnRaw, Cfg := cfg, NeutralXMem := nx, NeutralYMem := ny);
home(DeadmanArmed := joy.DeadmanArmed, JoystickDeflected := NOT joy.AtNeutralXY, JoystickPull := joy.AxisCmdY.DirectionPositive, JoystickPush := joy.AxisCmdY.DirectionNegative, BtnValidation := bench.Operator.JoyBtnRaw);
IF bench.Operator.JoyBtnRaw AND NOT previousButton THEN buttonEdges := buttonEdges + 1; END_IF; previousButton := bench.Operator.JoyBtnRaw;
ADVANCE_TIME(10000000);
bench(RawPosM1 := raw1, RawPosM2 := raw2);
joy(RawX := bench.Operator.JoyXRaw_ANA1, RawY := bench.Operator.JoyYRaw_ANA2, RawButton := bench.Operator.JoyBtnRaw, Cfg := cfg, NeutralXMem := nx, NeutralYMem := ny);
home(DeadmanArmed := joy.DeadmanArmed, JoystickDeflected := NOT joy.AtNeutralXY, JoystickPull := joy.AxisCmdY.DirectionPositive, JoystickPush := joy.AxisCmdY.DirectionNegative, BtnValidation := bench.Operator.JoyBtnRaw);
IF bench.Operator.JoyBtnRaw AND NOT previousButton THEN buttonEdges := buttonEdges + 1; END_IF; previousButton := bench.Operator.JoyBtnRaw;
ADVANCE_TIME(10000000);
bench(RawPosM1 := raw1, RawPosM2 := raw2);
joy(RawX := bench.Operator.JoyXRaw_ANA1, RawY := bench.Operator.JoyYRaw_ANA2, RawButton := bench.Operator.JoyBtnRaw, Cfg := cfg, NeutralXMem := nx, NeutralYMem := ny);
home(DeadmanArmed := joy.DeadmanArmed, JoystickDeflected := NOT joy.AtNeutralXY, JoystickPull := joy.AxisCmdY.DirectionPositive, JoystickPush := joy.AxisCmdY.DirectionNegative, BtnValidation := bench.Operator.JoyBtnRaw);
IF bench.Operator.JoyBtnRaw AND NOT previousButton THEN buttonEdges := buttonEdges + 1; END_IF; previousButton := bench.Operator.JoyBtnRaw;
ADVANCE_TIME(10000000);
bench(RawPosM1 := raw1, RawPosM2 := raw2);
joy(RawX := bench.Operator.JoyXRaw_ANA1, RawY := bench.Operator.JoyYRaw_ANA2, RawButton := bench.Operator.JoyBtnRaw, Cfg := cfg, NeutralXMem := nx, NeutralYMem := ny);
home(DeadmanArmed := joy.DeadmanArmed, JoystickDeflected := NOT joy.AtNeutralXY, JoystickPull := joy.AxisCmdY.DirectionPositive, JoystickPush := joy.AxisCmdY.DirectionNegative, BtnValidation := bench.Operator.JoyBtnRaw);
IF bench.Operator.JoyBtnRaw AND NOT previousButton THEN buttonEdges := buttonEdges + 1; END_IF; previousButton := bench.Operator.JoyBtnRaw;
ADVANCE_TIME(10000000);
bench(RawPosM1 := raw1, RawPosM2 := raw2);
joy(RawX := bench.Operator.JoyXRaw_ANA1, RawY := bench.Operator.JoyYRaw_ANA2, RawButton := bench.Operator.JoyBtnRaw, Cfg := cfg, NeutralXMem := nx, NeutralYMem := ny);
home(DeadmanArmed := joy.DeadmanArmed, JoystickDeflected := NOT joy.AtNeutralXY, JoystickPull := joy.AxisCmdY.DirectionPositive, JoystickPush := joy.AxisCmdY.DirectionNegative, BtnValidation := bench.Operator.JoyBtnRaw);
IF bench.Operator.JoyBtnRaw AND NOT previousButton THEN buttonEdges := buttonEdges + 1; END_IF; previousButton := bench.Operator.JoyBtnRaw;
ASSERT_FALSE(bench.Operator.JoyBtnRaw, 'Armement simule relache'); ASSERT_TRUE(joy.AxisCmdX.StartStop, 'Commande reelle active apres relachement'); ASSERT_TRUE(joy.DeadmanArmed, 'Armement reel conserve'); ASSERT_EQ(buttonEdges, 1, 'Un seul front brut');
bench.SimJoystickRight_Fwd_MAINT_Active := FALSE;
ADVANCE_TIME(10000000);
bench(RawPosM1 := raw1, RawPosM2 := raw2);
joy(RawX := bench.Operator.JoyXRaw_ANA1, RawY := bench.Operator.JoyYRaw_ANA2, RawButton := bench.Operator.JoyBtnRaw, Cfg := cfg, NeutralXMem := nx, NeutralYMem := ny);
home(DeadmanArmed := joy.DeadmanArmed, JoystickDeflected := NOT joy.AtNeutralXY, JoystickPull := joy.AxisCmdY.DirectionPositive, JoystickPush := joy.AxisCmdY.DirectionNegative, BtnValidation := bench.Operator.JoyBtnRaw);
IF bench.Operator.JoyBtnRaw AND NOT previousButton THEN buttonEdges := buttonEdges + 1; END_IF; previousButton := bench.Operator.JoyBtnRaw;
ADVANCE_TIME(10000000);
bench(RawPosM1 := raw1, RawPosM2 := raw2);
joy(RawX := bench.Operator.JoyXRaw_ANA1, RawY := bench.Operator.JoyYRaw_ANA2, RawButton := bench.Operator.JoyBtnRaw, Cfg := cfg, NeutralXMem := nx, NeutralYMem := ny);
home(DeadmanArmed := joy.DeadmanArmed, JoystickDeflected := NOT joy.AtNeutralXY, JoystickPull := joy.AxisCmdY.DirectionPositive, JoystickPush := joy.AxisCmdY.DirectionNegative, BtnValidation := bench.Operator.JoyBtnRaw);
IF bench.Operator.JoyBtnRaw AND NOT previousButton THEN buttonEdges := buttonEdges + 1; END_IF; previousButton := bench.Operator.JoyBtnRaw;
ADVANCE_TIME(10000000);
bench(RawPosM1 := raw1, RawPosM2 := raw2);
joy(RawX := bench.Operator.JoyXRaw_ANA1, RawY := bench.Operator.JoyYRaw_ANA2, RawButton := bench.Operator.JoyBtnRaw, Cfg := cfg, NeutralXMem := nx, NeutralYMem := ny);
home(DeadmanArmed := joy.DeadmanArmed, JoystickDeflected := NOT joy.AtNeutralXY, JoystickPull := joy.AxisCmdY.DirectionPositive, JoystickPush := joy.AxisCmdY.DirectionNegative, BtnValidation := bench.Operator.JoyBtnRaw);
IF bench.Operator.JoyBtnRaw AND NOT previousButton THEN buttonEdges := buttonEdges + 1; END_IF; previousButton := bench.Operator.JoyBtnRaw;
ADVANCE_TIME(10000000);
bench(RawPosM1 := raw1, RawPosM2 := raw2);
joy(RawX := bench.Operator.JoyXRaw_ANA1, RawY := bench.Operator.JoyYRaw_ANA2, RawButton := bench.Operator.JoyBtnRaw, Cfg := cfg, NeutralXMem := nx, NeutralYMem := ny);
home(DeadmanArmed := joy.DeadmanArmed, JoystickDeflected := NOT joy.AtNeutralXY, JoystickPull := joy.AxisCmdY.DirectionPositive, JoystickPush := joy.AxisCmdY.DirectionNegative, BtnValidation := bench.Operator.JoyBtnRaw);
IF bench.Operator.JoyBtnRaw AND NOT previousButton THEN buttonEdges := buttonEdges + 1; END_IF; previousButton := bench.Operator.JoyBtnRaw;
ADVANCE_TIME(10000000);
bench(RawPosM1 := raw1, RawPosM2 := raw2);
joy(RawX := bench.Operator.JoyXRaw_ANA1, RawY := bench.Operator.JoyYRaw_ANA2, RawButton := bench.Operator.JoyBtnRaw, Cfg := cfg, NeutralXMem := nx, NeutralYMem := ny);
home(DeadmanArmed := joy.DeadmanArmed, JoystickDeflected := NOT joy.AtNeutralXY, JoystickPull := joy.AxisCmdY.DirectionPositive, JoystickPush := joy.AxisCmdY.DirectionNegative, BtnValidation := bench.Operator.JoyBtnRaw);
IF bench.Operator.JoyBtnRaw AND NOT previousButton THEN buttonEdges := buttonEdges + 1; END_IF; previousButton := bench.Operator.JoyBtnRaw;
ADVANCE_TIME(10000000);
bench(RawPosM1 := raw1, RawPosM2 := raw2);
joy(RawX := bench.Operator.JoyXRaw_ANA1, RawY := bench.Operator.JoyYRaw_ANA2, RawButton := bench.Operator.JoyBtnRaw, Cfg := cfg, NeutralXMem := nx, NeutralYMem := ny);
home(DeadmanArmed := joy.DeadmanArmed, JoystickDeflected := NOT joy.AtNeutralXY, JoystickPull := joy.AxisCmdY.DirectionPositive, JoystickPush := joy.AxisCmdY.DirectionNegative, BtnValidation := bench.Operator.JoyBtnRaw);
IF bench.Operator.JoyBtnRaw AND NOT previousButton THEN buttonEdges := buttonEdges + 1; END_IF; previousButton := bench.Operator.JoyBtnRaw;
ADVANCE_TIME(10000000);
bench(RawPosM1 := raw1, RawPosM2 := raw2);
joy(RawX := bench.Operator.JoyXRaw_ANA1, RawY := bench.Operator.JoyYRaw_ANA2, RawButton := bench.Operator.JoyBtnRaw, Cfg := cfg, NeutralXMem := nx, NeutralYMem := ny);
home(DeadmanArmed := joy.DeadmanArmed, JoystickDeflected := NOT joy.AtNeutralXY, JoystickPull := joy.AxisCmdY.DirectionPositive, JoystickPush := joy.AxisCmdY.DirectionNegative, BtnValidation := bench.Operator.JoyBtnRaw);
IF bench.Operator.JoyBtnRaw AND NOT previousButton THEN buttonEdges := buttonEdges + 1; END_IF; previousButton := bench.Operator.JoyBtnRaw;
ADVANCE_TIME(10000000);
bench(RawPosM1 := raw1, RawPosM2 := raw2);
joy(RawX := bench.Operator.JoyXRaw_ANA1, RawY := bench.Operator.JoyYRaw_ANA2, RawButton := bench.Operator.JoyBtnRaw, Cfg := cfg, NeutralXMem := nx, NeutralYMem := ny);
home(DeadmanArmed := joy.DeadmanArmed, JoystickDeflected := NOT joy.AtNeutralXY, JoystickPull := joy.AxisCmdY.DirectionPositive, JoystickPush := joy.AxisCmdY.DirectionNegative, BtnValidation := bench.Operator.JoyBtnRaw);
IF bench.Operator.JoyBtnRaw AND NOT previousButton THEN buttonEdges := buttonEdges + 1; END_IF; previousButton := bench.Operator.JoyBtnRaw;
ADVANCE_TIME(10000000);
bench(RawPosM1 := raw1, RawPosM2 := raw2);
joy(RawX := bench.Operator.JoyXRaw_ANA1, RawY := bench.Operator.JoyYRaw_ANA2, RawButton := bench.Operator.JoyBtnRaw, Cfg := cfg, NeutralXMem := nx, NeutralYMem := ny);
home(DeadmanArmed := joy.DeadmanArmed, JoystickDeflected := NOT joy.AtNeutralXY, JoystickPull := joy.AxisCmdY.DirectionPositive, JoystickPush := joy.AxisCmdY.DirectionNegative, BtnValidation := bench.Operator.JoyBtnRaw);
IF bench.Operator.JoyBtnRaw AND NOT previousButton THEN buttonEdges := buttonEdges + 1; END_IF; previousButton := bench.Operator.JoyBtnRaw;
ADVANCE_TIME(10000000);
bench(RawPosM1 := raw1, RawPosM2 := raw2);
joy(RawX := bench.Operator.JoyXRaw_ANA1, RawY := bench.Operator.JoyYRaw_ANA2, RawButton := bench.Operator.JoyBtnRaw, Cfg := cfg, NeutralXMem := nx, NeutralYMem := ny);
home(DeadmanArmed := joy.DeadmanArmed, JoystickDeflected := NOT joy.AtNeutralXY, JoystickPull := joy.AxisCmdY.DirectionPositive, JoystickPush := joy.AxisCmdY.DirectionNegative, BtnValidation := bench.Operator.JoyBtnRaw);
IF bench.Operator.JoyBtnRaw AND NOT previousButton THEN buttonEdges := buttonEdges + 1; END_IF; previousButton := bench.Operator.JoyBtnRaw;
ADVANCE_TIME(10000000);
bench(RawPosM1 := raw1, RawPosM2 := raw2);
joy(RawX := bench.Operator.JoyXRaw_ANA1, RawY := bench.Operator.JoyYRaw_ANA2, RawButton := bench.Operator.JoyBtnRaw, Cfg := cfg, NeutralXMem := nx, NeutralYMem := ny);
home(DeadmanArmed := joy.DeadmanArmed, JoystickDeflected := NOT joy.AtNeutralXY, JoystickPull := joy.AxisCmdY.DirectionPositive, JoystickPush := joy.AxisCmdY.DirectionNegative, BtnValidation := bench.Operator.JoyBtnRaw);
IF bench.Operator.JoyBtnRaw AND NOT previousButton THEN buttonEdges := buttonEdges + 1; END_IF; previousButton := bench.Operator.JoyBtnRaw;
ADVANCE_TIME(10000000);
bench(RawPosM1 := raw1, RawPosM2 := raw2);
joy(RawX := bench.Operator.JoyXRaw_ANA1, RawY := bench.Operator.JoyYRaw_ANA2, RawButton := bench.Operator.JoyBtnRaw, Cfg := cfg, NeutralXMem := nx, NeutralYMem := ny);
home(DeadmanArmed := joy.DeadmanArmed, JoystickDeflected := NOT joy.AtNeutralXY, JoystickPull := joy.AxisCmdY.DirectionPositive, JoystickPush := joy.AxisCmdY.DirectionNegative, BtnValidation := bench.Operator.JoyBtnRaw);
IF bench.Operator.JoyBtnRaw AND NOT previousButton THEN buttonEdges := buttonEdges + 1; END_IF; previousButton := bench.Operator.JoyBtnRaw;
ADVANCE_TIME(10000000);
bench(RawPosM1 := raw1, RawPosM2 := raw2);
joy(RawX := bench.Operator.JoyXRaw_ANA1, RawY := bench.Operator.JoyYRaw_ANA2, RawButton := bench.Operator.JoyBtnRaw, Cfg := cfg, NeutralXMem := nx, NeutralYMem := ny);
home(DeadmanArmed := joy.DeadmanArmed, JoystickDeflected := NOT joy.AtNeutralXY, JoystickPull := joy.AxisCmdY.DirectionPositive, JoystickPush := joy.AxisCmdY.DirectionNegative, BtnValidation := bench.Operator.JoyBtnRaw);
IF bench.Operator.JoyBtnRaw AND NOT previousButton THEN buttonEdges := buttonEdges + 1; END_IF; previousButton := bench.Operator.JoyBtnRaw;
ADVANCE_TIME(10000000);
bench(RawPosM1 := raw1, RawPosM2 := raw2);
joy(RawX := bench.Operator.JoyXRaw_ANA1, RawY := bench.Operator.JoyYRaw_ANA2, RawButton := bench.Operator.JoyBtnRaw, Cfg := cfg, NeutralXMem := nx, NeutralYMem := ny);
home(DeadmanArmed := joy.DeadmanArmed, JoystickDeflected := NOT joy.AtNeutralXY, JoystickPull := joy.AxisCmdY.DirectionPositive, JoystickPush := joy.AxisCmdY.DirectionNegative, BtnValidation := bench.Operator.JoyBtnRaw);
IF bench.Operator.JoyBtnRaw AND NOT previousButton THEN buttonEdges := buttonEdges + 1; END_IF; previousButton := bench.Operator.JoyBtnRaw;
ADVANCE_TIME(10000000);
bench(RawPosM1 := raw1, RawPosM2 := raw2);
joy(RawX := bench.Operator.JoyXRaw_ANA1, RawY := bench.Operator.JoyYRaw_ANA2, RawButton := bench.Operator.JoyBtnRaw, Cfg := cfg, NeutralXMem := nx, NeutralYMem := ny);
home(DeadmanArmed := joy.DeadmanArmed, JoystickDeflected := NOT joy.AtNeutralXY, JoystickPull := joy.AxisCmdY.DirectionPositive, JoystickPush := joy.AxisCmdY.DirectionNegative, BtnValidation := bench.Operator.JoyBtnRaw);
IF bench.Operator.JoyBtnRaw AND NOT previousButton THEN buttonEdges := buttonEdges + 1; END_IF; previousButton := bench.Operator.JoyBtnRaw;
ADVANCE_TIME(10000000);
bench(RawPosM1 := raw1, RawPosM2 := raw2);
joy(RawX := bench.Operator.JoyXRaw_ANA1, RawY := bench.Operator.JoyYRaw_ANA2, RawButton := bench.Operator.JoyBtnRaw, Cfg := cfg, NeutralXMem := nx, NeutralYMem := ny);
home(DeadmanArmed := joy.DeadmanArmed, JoystickDeflected := NOT joy.AtNeutralXY, JoystickPull := joy.AxisCmdY.DirectionPositive, JoystickPush := joy.AxisCmdY.DirectionNegative, BtnValidation := bench.Operator.JoyBtnRaw);
IF bench.Operator.JoyBtnRaw AND NOT previousButton THEN buttonEdges := buttonEdges + 1; END_IF; previousButton := bench.Operator.JoyBtnRaw;
ADVANCE_TIME(10000000);
bench(RawPosM1 := raw1, RawPosM2 := raw2);
joy(RawX := bench.Operator.JoyXRaw_ANA1, RawY := bench.Operator.JoyYRaw_ANA2, RawButton := bench.Operator.JoyBtnRaw, Cfg := cfg, NeutralXMem := nx, NeutralYMem := ny);
home(DeadmanArmed := joy.DeadmanArmed, JoystickDeflected := NOT joy.AtNeutralXY, JoystickPull := joy.AxisCmdY.DirectionPositive, JoystickPush := joy.AxisCmdY.DirectionNegative, BtnValidation := bench.Operator.JoyBtnRaw);
IF bench.Operator.JoyBtnRaw AND NOT previousButton THEN buttonEdges := buttonEdges + 1; END_IF; previousButton := bench.Operator.JoyBtnRaw;
ADVANCE_TIME(10000000);
bench(RawPosM1 := raw1, RawPosM2 := raw2);
joy(RawX := bench.Operator.JoyXRaw_ANA1, RawY := bench.Operator.JoyYRaw_ANA2, RawButton := bench.Operator.JoyBtnRaw, Cfg := cfg, NeutralXMem := nx, NeutralYMem := ny);
home(DeadmanArmed := joy.DeadmanArmed, JoystickDeflected := NOT joy.AtNeutralXY, JoystickPull := joy.AxisCmdY.DirectionPositive, JoystickPush := joy.AxisCmdY.DirectionNegative, BtnValidation := bench.Operator.JoyBtnRaw);
IF bench.Operator.JoyBtnRaw AND NOT previousButton THEN buttonEdges := buttonEdges + 1; END_IF; previousButton := bench.Operator.JoyBtnRaw;
ADVANCE_TIME(10000000);
bench(RawPosM1 := raw1, RawPosM2 := raw2);
joy(RawX := bench.Operator.JoyXRaw_ANA1, RawY := bench.Operator.JoyYRaw_ANA2, RawButton := bench.Operator.JoyBtnRaw, Cfg := cfg, NeutralXMem := nx, NeutralYMem := ny);
home(DeadmanArmed := joy.DeadmanArmed, JoystickDeflected := NOT joy.AtNeutralXY, JoystickPull := joy.AxisCmdY.DirectionPositive, JoystickPush := joy.AxisCmdY.DirectionNegative, BtnValidation := bench.Operator.JoyBtnRaw);
IF bench.Operator.JoyBtnRaw AND NOT previousButton THEN buttonEdges := buttonEdges + 1; END_IF; previousButton := bench.Operator.JoyBtnRaw;
ADVANCE_TIME(10000000);
bench(RawPosM1 := raw1, RawPosM2 := raw2);
joy(RawX := bench.Operator.JoyXRaw_ANA1, RawY := bench.Operator.JoyYRaw_ANA2, RawButton := bench.Operator.JoyBtnRaw, Cfg := cfg, NeutralXMem := nx, NeutralYMem := ny);
home(DeadmanArmed := joy.DeadmanArmed, JoystickDeflected := NOT joy.AtNeutralXY, JoystickPull := joy.AxisCmdY.DirectionPositive, JoystickPush := joy.AxisCmdY.DirectionNegative, BtnValidation := bench.Operator.JoyBtnRaw);
IF bench.Operator.JoyBtnRaw AND NOT previousButton THEN buttonEdges := buttonEdges + 1; END_IF; previousButton := bench.Operator.JoyBtnRaw;
ADVANCE_TIME(10000000);
bench(RawPosM1 := raw1, RawPosM2 := raw2);
joy(RawX := bench.Operator.JoyXRaw_ANA1, RawY := bench.Operator.JoyYRaw_ANA2, RawButton := bench.Operator.JoyBtnRaw, Cfg := cfg, NeutralXMem := nx, NeutralYMem := ny);
home(DeadmanArmed := joy.DeadmanArmed, JoystickDeflected := NOT joy.AtNeutralXY, JoystickPull := joy.AxisCmdY.DirectionPositive, JoystickPush := joy.AxisCmdY.DirectionNegative, BtnValidation := bench.Operator.JoyBtnRaw);
IF bench.Operator.JoyBtnRaw AND NOT previousButton THEN buttonEdges := buttonEdges + 1; END_IF; previousButton := bench.Operator.JoyBtnRaw;
ADVANCE_TIME(10000000);
bench(RawPosM1 := raw1, RawPosM2 := raw2);
joy(RawX := bench.Operator.JoyXRaw_ANA1, RawY := bench.Operator.JoyYRaw_ANA2, RawButton := bench.Operator.JoyBtnRaw, Cfg := cfg, NeutralXMem := nx, NeutralYMem := ny);
home(DeadmanArmed := joy.DeadmanArmed, JoystickDeflected := NOT joy.AtNeutralXY, JoystickPull := joy.AxisCmdY.DirectionPositive, JoystickPush := joy.AxisCmdY.DirectionNegative, BtnValidation := bench.Operator.JoyBtnRaw);
IF bench.Operator.JoyBtnRaw AND NOT previousButton THEN buttonEdges := buttonEdges + 1; END_IF; previousButton := bench.Operator.JoyBtnRaw;
ADVANCE_TIME(10000000);
bench(RawPosM1 := raw1, RawPosM2 := raw2);
joy(RawX := bench.Operator.JoyXRaw_ANA1, RawY := bench.Operator.JoyYRaw_ANA2, RawButton := bench.Operator.JoyBtnRaw, Cfg := cfg, NeutralXMem := nx, NeutralYMem := ny);
home(DeadmanArmed := joy.DeadmanArmed, JoystickDeflected := NOT joy.AtNeutralXY, JoystickPull := joy.AxisCmdY.DirectionPositive, JoystickPush := joy.AxisCmdY.DirectionNegative, BtnValidation := bench.Operator.JoyBtnRaw);
IF bench.Operator.JoyBtnRaw AND NOT previousButton THEN buttonEdges := buttonEdges + 1; END_IF; previousButton := bench.Operator.JoyBtnRaw;
ADVANCE_TIME(10000000);
bench(RawPosM1 := raw1, RawPosM2 := raw2);
joy(RawX := bench.Operator.JoyXRaw_ANA1, RawY := bench.Operator.JoyYRaw_ANA2, RawButton := bench.Operator.JoyBtnRaw, Cfg := cfg, NeutralXMem := nx, NeutralYMem := ny);
home(DeadmanArmed := joy.DeadmanArmed, JoystickDeflected := NOT joy.AtNeutralXY, JoystickPull := joy.AxisCmdY.DirectionPositive, JoystickPush := joy.AxisCmdY.DirectionNegative, BtnValidation := bench.Operator.JoyBtnRaw);
IF bench.Operator.JoyBtnRaw AND NOT previousButton THEN buttonEdges := buttonEdges + 1; END_IF; previousButton := bench.Operator.JoyBtnRaw;
ADVANCE_TIME(10000000);
bench(RawPosM1 := raw1, RawPosM2 := raw2);
joy(RawX := bench.Operator.JoyXRaw_ANA1, RawY := bench.Operator.JoyYRaw_ANA2, RawButton := bench.Operator.JoyBtnRaw, Cfg := cfg, NeutralXMem := nx, NeutralYMem := ny);
home(DeadmanArmed := joy.DeadmanArmed, JoystickDeflected := NOT joy.AtNeutralXY, JoystickPull := joy.AxisCmdY.DirectionPositive, JoystickPush := joy.AxisCmdY.DirectionNegative, BtnValidation := bench.Operator.JoyBtnRaw);
IF bench.Operator.JoyBtnRaw AND NOT previousButton THEN buttonEdges := buttonEdges + 1; END_IF; previousButton := bench.Operator.JoyBtnRaw;
ASSERT_TRUE(joy.AtNeutralXY, 'Retour neutre'); ASSERT_FALSE(joy.AxisCmdX.StartStop, 'Commande nulle au neutre'); ASSERT_TRUE(joy.DeadmanArmed, 'Grace conserve armement sur geste court');
bench.SimJoystickLeft_Rev_TREMIE_Active := TRUE;
ADVANCE_TIME(10000000);
bench(RawPosM1 := raw1, RawPosM2 := raw2);
joy(RawX := bench.Operator.JoyXRaw_ANA1, RawY := bench.Operator.JoyYRaw_ANA2, RawButton := bench.Operator.JoyBtnRaw, Cfg := cfg, NeutralXMem := nx, NeutralYMem := ny);
home(DeadmanArmed := joy.DeadmanArmed, JoystickDeflected := NOT joy.AtNeutralXY, JoystickPull := joy.AxisCmdY.DirectionPositive, JoystickPush := joy.AxisCmdY.DirectionNegative, BtnValidation := bench.Operator.JoyBtnRaw);
IF bench.Operator.JoyBtnRaw AND NOT previousButton THEN buttonEdges := buttonEdges + 1; END_IF; previousButton := bench.Operator.JoyBtnRaw;
ADVANCE_TIME(10000000);
bench(RawPosM1 := raw1, RawPosM2 := raw2);
joy(RawX := bench.Operator.JoyXRaw_ANA1, RawY := bench.Operator.JoyYRaw_ANA2, RawButton := bench.Operator.JoyBtnRaw, Cfg := cfg, NeutralXMem := nx, NeutralYMem := ny);
home(DeadmanArmed := joy.DeadmanArmed, JoystickDeflected := NOT joy.AtNeutralXY, JoystickPull := joy.AxisCmdY.DirectionPositive, JoystickPush := joy.AxisCmdY.DirectionNegative, BtnValidation := bench.Operator.JoyBtnRaw);
IF bench.Operator.JoyBtnRaw AND NOT previousButton THEN buttonEdges := buttonEdges + 1; END_IF; previousButton := bench.Operator.JoyBtnRaw;
ADVANCE_TIME(10000000);
bench(RawPosM1 := raw1, RawPosM2 := raw2);
joy(RawX := bench.Operator.JoyXRaw_ANA1, RawY := bench.Operator.JoyYRaw_ANA2, RawButton := bench.Operator.JoyBtnRaw, Cfg := cfg, NeutralXMem := nx, NeutralYMem := ny);
home(DeadmanArmed := joy.DeadmanArmed, JoystickDeflected := NOT joy.AtNeutralXY, JoystickPull := joy.AxisCmdY.DirectionPositive, JoystickPush := joy.AxisCmdY.DirectionNegative, BtnValidation := bench.Operator.JoyBtnRaw);
IF bench.Operator.JoyBtnRaw AND NOT previousButton THEN buttonEdges := buttonEdges + 1; END_IF; previousButton := bench.Operator.JoyBtnRaw;
ADVANCE_TIME(10000000);
bench(RawPosM1 := raw1, RawPosM2 := raw2);
joy(RawX := bench.Operator.JoyXRaw_ANA1, RawY := bench.Operator.JoyYRaw_ANA2, RawButton := bench.Operator.JoyBtnRaw, Cfg := cfg, NeutralXMem := nx, NeutralYMem := ny);
home(DeadmanArmed := joy.DeadmanArmed, JoystickDeflected := NOT joy.AtNeutralXY, JoystickPull := joy.AxisCmdY.DirectionPositive, JoystickPush := joy.AxisCmdY.DirectionNegative, BtnValidation := bench.Operator.JoyBtnRaw);
IF bench.Operator.JoyBtnRaw AND NOT previousButton THEN buttonEdges := buttonEdges + 1; END_IF; previousButton := bench.Operator.JoyBtnRaw;
ADVANCE_TIME(10000000);
bench(RawPosM1 := raw1, RawPosM2 := raw2);
joy(RawX := bench.Operator.JoyXRaw_ANA1, RawY := bench.Operator.JoyYRaw_ANA2, RawButton := bench.Operator.JoyBtnRaw, Cfg := cfg, NeutralXMem := nx, NeutralYMem := ny);
home(DeadmanArmed := joy.DeadmanArmed, JoystickDeflected := NOT joy.AtNeutralXY, JoystickPull := joy.AxisCmdY.DirectionPositive, JoystickPush := joy.AxisCmdY.DirectionNegative, BtnValidation := bench.Operator.JoyBtnRaw);
IF bench.Operator.JoyBtnRaw AND NOT previousButton THEN buttonEdges := buttonEdges + 1; END_IF; previousButton := bench.Operator.JoyBtnRaw;
ADVANCE_TIME(10000000);
bench(RawPosM1 := raw1, RawPosM2 := raw2);
joy(RawX := bench.Operator.JoyXRaw_ANA1, RawY := bench.Operator.JoyYRaw_ANA2, RawButton := bench.Operator.JoyBtnRaw, Cfg := cfg, NeutralXMem := nx, NeutralYMem := ny);
home(DeadmanArmed := joy.DeadmanArmed, JoystickDeflected := NOT joy.AtNeutralXY, JoystickPull := joy.AxisCmdY.DirectionPositive, JoystickPush := joy.AxisCmdY.DirectionNegative, BtnValidation := bench.Operator.JoyBtnRaw);
IF bench.Operator.JoyBtnRaw AND NOT previousButton THEN buttonEdges := buttonEdges + 1; END_IF; previousButton := bench.Operator.JoyBtnRaw;
ADVANCE_TIME(10000000);
bench(RawPosM1 := raw1, RawPosM2 := raw2);
joy(RawX := bench.Operator.JoyXRaw_ANA1, RawY := bench.Operator.JoyYRaw_ANA2, RawButton := bench.Operator.JoyBtnRaw, Cfg := cfg, NeutralXMem := nx, NeutralYMem := ny);
home(DeadmanArmed := joy.DeadmanArmed, JoystickDeflected := NOT joy.AtNeutralXY, JoystickPull := joy.AxisCmdY.DirectionPositive, JoystickPush := joy.AxisCmdY.DirectionNegative, BtnValidation := bench.Operator.JoyBtnRaw);
IF bench.Operator.JoyBtnRaw AND NOT previousButton THEN buttonEdges := buttonEdges + 1; END_IF; previousButton := bench.Operator.JoyBtnRaw;
ADVANCE_TIME(10000000);
bench(RawPosM1 := raw1, RawPosM2 := raw2);
joy(RawX := bench.Operator.JoyXRaw_ANA1, RawY := bench.Operator.JoyYRaw_ANA2, RawButton := bench.Operator.JoyBtnRaw, Cfg := cfg, NeutralXMem := nx, NeutralYMem := ny);
home(DeadmanArmed := joy.DeadmanArmed, JoystickDeflected := NOT joy.AtNeutralXY, JoystickPull := joy.AxisCmdY.DirectionPositive, JoystickPush := joy.AxisCmdY.DirectionNegative, BtnValidation := bench.Operator.JoyBtnRaw);
IF bench.Operator.JoyBtnRaw AND NOT previousButton THEN buttonEdges := buttonEdges + 1; END_IF; previousButton := bench.Operator.JoyBtnRaw;
ADVANCE_TIME(10000000);
bench(RawPosM1 := raw1, RawPosM2 := raw2);
joy(RawX := bench.Operator.JoyXRaw_ANA1, RawY := bench.Operator.JoyYRaw_ANA2, RawButton := bench.Operator.JoyBtnRaw, Cfg := cfg, NeutralXMem := nx, NeutralYMem := ny);
home(DeadmanArmed := joy.DeadmanArmed, JoystickDeflected := NOT joy.AtNeutralXY, JoystickPull := joy.AxisCmdY.DirectionPositive, JoystickPush := joy.AxisCmdY.DirectionNegative, BtnValidation := bench.Operator.JoyBtnRaw);
IF bench.Operator.JoyBtnRaw AND NOT previousButton THEN buttonEdges := buttonEdges + 1; END_IF; previousButton := bench.Operator.JoyBtnRaw;
ADVANCE_TIME(10000000);
bench(RawPosM1 := raw1, RawPosM2 := raw2);
joy(RawX := bench.Operator.JoyXRaw_ANA1, RawY := bench.Operator.JoyYRaw_ANA2, RawButton := bench.Operator.JoyBtnRaw, Cfg := cfg, NeutralXMem := nx, NeutralYMem := ny);
home(DeadmanArmed := joy.DeadmanArmed, JoystickDeflected := NOT joy.AtNeutralXY, JoystickPull := joy.AxisCmdY.DirectionPositive, JoystickPush := joy.AxisCmdY.DirectionNegative, BtnValidation := bench.Operator.JoyBtnRaw);
IF bench.Operator.JoyBtnRaw AND NOT previousButton THEN buttonEdges := buttonEdges + 1; END_IF; previousButton := bench.Operator.JoyBtnRaw;
ADVANCE_TIME(10000000);
bench(RawPosM1 := raw1, RawPosM2 := raw2);
joy(RawX := bench.Operator.JoyXRaw_ANA1, RawY := bench.Operator.JoyYRaw_ANA2, RawButton := bench.Operator.JoyBtnRaw, Cfg := cfg, NeutralXMem := nx, NeutralYMem := ny);
home(DeadmanArmed := joy.DeadmanArmed, JoystickDeflected := NOT joy.AtNeutralXY, JoystickPull := joy.AxisCmdY.DirectionPositive, JoystickPush := joy.AxisCmdY.DirectionNegative, BtnValidation := bench.Operator.JoyBtnRaw);
IF bench.Operator.JoyBtnRaw AND NOT previousButton THEN buttonEdges := buttonEdges + 1; END_IF; previousButton := bench.Operator.JoyBtnRaw;
ADVANCE_TIME(10000000);
bench(RawPosM1 := raw1, RawPosM2 := raw2);
joy(RawX := bench.Operator.JoyXRaw_ANA1, RawY := bench.Operator.JoyYRaw_ANA2, RawButton := bench.Operator.JoyBtnRaw, Cfg := cfg, NeutralXMem := nx, NeutralYMem := ny);
home(DeadmanArmed := joy.DeadmanArmed, JoystickDeflected := NOT joy.AtNeutralXY, JoystickPull := joy.AxisCmdY.DirectionPositive, JoystickPush := joy.AxisCmdY.DirectionNegative, BtnValidation := bench.Operator.JoyBtnRaw);
IF bench.Operator.JoyBtnRaw AND NOT previousButton THEN buttonEdges := buttonEdges + 1; END_IF; previousButton := bench.Operator.JoyBtnRaw;
ADVANCE_TIME(10000000);
bench(RawPosM1 := raw1, RawPosM2 := raw2);
joy(RawX := bench.Operator.JoyXRaw_ANA1, RawY := bench.Operator.JoyYRaw_ANA2, RawButton := bench.Operator.JoyBtnRaw, Cfg := cfg, NeutralXMem := nx, NeutralYMem := ny);
home(DeadmanArmed := joy.DeadmanArmed, JoystickDeflected := NOT joy.AtNeutralXY, JoystickPull := joy.AxisCmdY.DirectionPositive, JoystickPush := joy.AxisCmdY.DirectionNegative, BtnValidation := bench.Operator.JoyBtnRaw);
IF bench.Operator.JoyBtnRaw AND NOT previousButton THEN buttonEdges := buttonEdges + 1; END_IF; previousButton := bench.Operator.JoyBtnRaw;
ADVANCE_TIME(10000000);
bench(RawPosM1 := raw1, RawPosM2 := raw2);
joy(RawX := bench.Operator.JoyXRaw_ANA1, RawY := bench.Operator.JoyYRaw_ANA2, RawButton := bench.Operator.JoyBtnRaw, Cfg := cfg, NeutralXMem := nx, NeutralYMem := ny);
home(DeadmanArmed := joy.DeadmanArmed, JoystickDeflected := NOT joy.AtNeutralXY, JoystickPull := joy.AxisCmdY.DirectionPositive, JoystickPush := joy.AxisCmdY.DirectionNegative, BtnValidation := bench.Operator.JoyBtnRaw);
IF bench.Operator.JoyBtnRaw AND NOT previousButton THEN buttonEdges := buttonEdges + 1; END_IF; previousButton := bench.Operator.JoyBtnRaw;
ADVANCE_TIME(10000000);
bench(RawPosM1 := raw1, RawPosM2 := raw2);
joy(RawX := bench.Operator.JoyXRaw_ANA1, RawY := bench.Operator.JoyYRaw_ANA2, RawButton := bench.Operator.JoyBtnRaw, Cfg := cfg, NeutralXMem := nx, NeutralYMem := ny);
home(DeadmanArmed := joy.DeadmanArmed, JoystickDeflected := NOT joy.AtNeutralXY, JoystickPull := joy.AxisCmdY.DirectionPositive, JoystickPush := joy.AxisCmdY.DirectionNegative, BtnValidation := bench.Operator.JoyBtnRaw);
IF bench.Operator.JoyBtnRaw AND NOT previousButton THEN buttonEdges := buttonEdges + 1; END_IF; previousButton := bench.Operator.JoyBtnRaw;
ADVANCE_TIME(10000000);
bench(RawPosM1 := raw1, RawPosM2 := raw2);
joy(RawX := bench.Operator.JoyXRaw_ANA1, RawY := bench.Operator.JoyYRaw_ANA2, RawButton := bench.Operator.JoyBtnRaw, Cfg := cfg, NeutralXMem := nx, NeutralYMem := ny);
home(DeadmanArmed := joy.DeadmanArmed, JoystickDeflected := NOT joy.AtNeutralXY, JoystickPull := joy.AxisCmdY.DirectionPositive, JoystickPush := joy.AxisCmdY.DirectionNegative, BtnValidation := bench.Operator.JoyBtnRaw);
IF bench.Operator.JoyBtnRaw AND NOT previousButton THEN buttonEdges := buttonEdges + 1; END_IF; previousButton := bench.Operator.JoyBtnRaw;
ADVANCE_TIME(10000000);
bench(RawPosM1 := raw1, RawPosM2 := raw2);
joy(RawX := bench.Operator.JoyXRaw_ANA1, RawY := bench.Operator.JoyYRaw_ANA2, RawButton := bench.Operator.JoyBtnRaw, Cfg := cfg, NeutralXMem := nx, NeutralYMem := ny);
home(DeadmanArmed := joy.DeadmanArmed, JoystickDeflected := NOT joy.AtNeutralXY, JoystickPull := joy.AxisCmdY.DirectionPositive, JoystickPush := joy.AxisCmdY.DirectionNegative, BtnValidation := bench.Operator.JoyBtnRaw);
IF bench.Operator.JoyBtnRaw AND NOT previousButton THEN buttonEdges := buttonEdges + 1; END_IF; previousButton := bench.Operator.JoyBtnRaw;
ADVANCE_TIME(10000000);
bench(RawPosM1 := raw1, RawPosM2 := raw2);
joy(RawX := bench.Operator.JoyXRaw_ANA1, RawY := bench.Operator.JoyYRaw_ANA2, RawButton := bench.Operator.JoyBtnRaw, Cfg := cfg, NeutralXMem := nx, NeutralYMem := ny);
home(DeadmanArmed := joy.DeadmanArmed, JoystickDeflected := NOT joy.AtNeutralXY, JoystickPull := joy.AxisCmdY.DirectionPositive, JoystickPush := joy.AxisCmdY.DirectionNegative, BtnValidation := bench.Operator.JoyBtnRaw);
IF bench.Operator.JoyBtnRaw AND NOT previousButton THEN buttonEdges := buttonEdges + 1; END_IF; previousButton := bench.Operator.JoyBtnRaw;
ADVANCE_TIME(10000000);
bench(RawPosM1 := raw1, RawPosM2 := raw2);
joy(RawX := bench.Operator.JoyXRaw_ANA1, RawY := bench.Operator.JoyYRaw_ANA2, RawButton := bench.Operator.JoyBtnRaw, Cfg := cfg, NeutralXMem := nx, NeutralYMem := ny);
home(DeadmanArmed := joy.DeadmanArmed, JoystickDeflected := NOT joy.AtNeutralXY, JoystickPull := joy.AxisCmdY.DirectionPositive, JoystickPush := joy.AxisCmdY.DirectionNegative, BtnValidation := bench.Operator.JoyBtnRaw);
IF bench.Operator.JoyBtnRaw AND NOT previousButton THEN buttonEdges := buttonEdges + 1; END_IF; previousButton := bench.Operator.JoyBtnRaw;
ADVANCE_TIME(10000000);
bench(RawPosM1 := raw1, RawPosM2 := raw2);
joy(RawX := bench.Operator.JoyXRaw_ANA1, RawY := bench.Operator.JoyYRaw_ANA2, RawButton := bench.Operator.JoyBtnRaw, Cfg := cfg, NeutralXMem := nx, NeutralYMem := ny);
home(DeadmanArmed := joy.DeadmanArmed, JoystickDeflected := NOT joy.AtNeutralXY, JoystickPull := joy.AxisCmdY.DirectionPositive, JoystickPush := joy.AxisCmdY.DirectionNegative, BtnValidation := bench.Operator.JoyBtnRaw);
IF bench.Operator.JoyBtnRaw AND NOT previousButton THEN buttonEdges := buttonEdges + 1; END_IF; previousButton := bench.Operator.JoyBtnRaw;
ADVANCE_TIME(10000000);
bench(RawPosM1 := raw1, RawPosM2 := raw2);
joy(RawX := bench.Operator.JoyXRaw_ANA1, RawY := bench.Operator.JoyYRaw_ANA2, RawButton := bench.Operator.JoyBtnRaw, Cfg := cfg, NeutralXMem := nx, NeutralYMem := ny);
home(DeadmanArmed := joy.DeadmanArmed, JoystickDeflected := NOT joy.AtNeutralXY, JoystickPull := joy.AxisCmdY.DirectionPositive, JoystickPush := joy.AxisCmdY.DirectionNegative, BtnValidation := bench.Operator.JoyBtnRaw);
IF bench.Operator.JoyBtnRaw AND NOT previousButton THEN buttonEdges := buttonEdges + 1; END_IF; previousButton := bench.Operator.JoyBtnRaw;
ADVANCE_TIME(10000000);
bench(RawPosM1 := raw1, RawPosM2 := raw2);
joy(RawX := bench.Operator.JoyXRaw_ANA1, RawY := bench.Operator.JoyYRaw_ANA2, RawButton := bench.Operator.JoyBtnRaw, Cfg := cfg, NeutralXMem := nx, NeutralYMem := ny);
home(DeadmanArmed := joy.DeadmanArmed, JoystickDeflected := NOT joy.AtNeutralXY, JoystickPull := joy.AxisCmdY.DirectionPositive, JoystickPush := joy.AxisCmdY.DirectionNegative, BtnValidation := bench.Operator.JoyBtnRaw);
IF bench.Operator.JoyBtnRaw AND NOT previousButton THEN buttonEdges := buttonEdges + 1; END_IF; previousButton := bench.Operator.JoyBtnRaw;
ADVANCE_TIME(10000000);
bench(RawPosM1 := raw1, RawPosM2 := raw2);
joy(RawX := bench.Operator.JoyXRaw_ANA1, RawY := bench.Operator.JoyYRaw_ANA2, RawButton := bench.Operator.JoyBtnRaw, Cfg := cfg, NeutralXMem := nx, NeutralYMem := ny);
home(DeadmanArmed := joy.DeadmanArmed, JoystickDeflected := NOT joy.AtNeutralXY, JoystickPull := joy.AxisCmdY.DirectionPositive, JoystickPush := joy.AxisCmdY.DirectionNegative, BtnValidation := bench.Operator.JoyBtnRaw);
IF bench.Operator.JoyBtnRaw AND NOT previousButton THEN buttonEdges := buttonEdges + 1; END_IF; previousButton := bench.Operator.JoyBtnRaw;
ADVANCE_TIME(10000000);
bench(RawPosM1 := raw1, RawPosM2 := raw2);
joy(RawX := bench.Operator.JoyXRaw_ANA1, RawY := bench.Operator.JoyYRaw_ANA2, RawButton := bench.Operator.JoyBtnRaw, Cfg := cfg, NeutralXMem := nx, NeutralYMem := ny);
home(DeadmanArmed := joy.DeadmanArmed, JoystickDeflected := NOT joy.AtNeutralXY, JoystickPull := joy.AxisCmdY.DirectionPositive, JoystickPush := joy.AxisCmdY.DirectionNegative, BtnValidation := bench.Operator.JoyBtnRaw);
IF bench.Operator.JoyBtnRaw AND NOT previousButton THEN buttonEdges := buttonEdges + 1; END_IF; previousButton := bench.Operator.JoyBtnRaw;
ADVANCE_TIME(10000000);
bench(RawPosM1 := raw1, RawPosM2 := raw2);
joy(RawX := bench.Operator.JoyXRaw_ANA1, RawY := bench.Operator.JoyYRaw_ANA2, RawButton := bench.Operator.JoyBtnRaw, Cfg := cfg, NeutralXMem := nx, NeutralYMem := ny);
home(DeadmanArmed := joy.DeadmanArmed, JoystickDeflected := NOT joy.AtNeutralXY, JoystickPull := joy.AxisCmdY.DirectionPositive, JoystickPush := joy.AxisCmdY.DirectionNegative, BtnValidation := bench.Operator.JoyBtnRaw);
IF bench.Operator.JoyBtnRaw AND NOT previousButton THEN buttonEdges := buttonEdges + 1; END_IF; previousButton := bench.Operator.JoyBtnRaw;
ADVANCE_TIME(10000000);
bench(RawPosM1 := raw1, RawPosM2 := raw2);
joy(RawX := bench.Operator.JoyXRaw_ANA1, RawY := bench.Operator.JoyYRaw_ANA2, RawButton := bench.Operator.JoyBtnRaw, Cfg := cfg, NeutralXMem := nx, NeutralYMem := ny);
home(DeadmanArmed := joy.DeadmanArmed, JoystickDeflected := NOT joy.AtNeutralXY, JoystickPull := joy.AxisCmdY.DirectionPositive, JoystickPush := joy.AxisCmdY.DirectionNegative, BtnValidation := bench.Operator.JoyBtnRaw);
IF bench.Operator.JoyBtnRaw AND NOT previousButton THEN buttonEdges := buttonEdges + 1; END_IF; previousButton := bench.Operator.JoyBtnRaw;
ADVANCE_TIME(10000000);
bench(RawPosM1 := raw1, RawPosM2 := raw2);
joy(RawX := bench.Operator.JoyXRaw_ANA1, RawY := bench.Operator.JoyYRaw_ANA2, RawButton := bench.Operator.JoyBtnRaw, Cfg := cfg, NeutralXMem := nx, NeutralYMem := ny);
home(DeadmanArmed := joy.DeadmanArmed, JoystickDeflected := NOT joy.AtNeutralXY, JoystickPull := joy.AxisCmdY.DirectionPositive, JoystickPush := joy.AxisCmdY.DirectionNegative, BtnValidation := bench.Operator.JoyBtnRaw);
IF bench.Operator.JoyBtnRaw AND NOT previousButton THEN buttonEdges := buttonEdges + 1; END_IF; previousButton := bench.Operator.JoyBtnRaw;
ADVANCE_TIME(10000000);
bench(RawPosM1 := raw1, RawPosM2 := raw2);
joy(RawX := bench.Operator.JoyXRaw_ANA1, RawY := bench.Operator.JoyYRaw_ANA2, RawButton := bench.Operator.JoyBtnRaw, Cfg := cfg, NeutralXMem := nx, NeutralYMem := ny);
home(DeadmanArmed := joy.DeadmanArmed, JoystickDeflected := NOT joy.AtNeutralXY, JoystickPull := joy.AxisCmdY.DirectionPositive, JoystickPush := joy.AxisCmdY.DirectionNegative, BtnValidation := bench.Operator.JoyBtnRaw);
IF bench.Operator.JoyBtnRaw AND NOT previousButton THEN buttonEdges := buttonEdges + 1; END_IF; previousButton := bench.Operator.JoyBtnRaw;
ADVANCE_TIME(10000000);
bench(RawPosM1 := raw1, RawPosM2 := raw2);
joy(RawX := bench.Operator.JoyXRaw_ANA1, RawY := bench.Operator.JoyYRaw_ANA2, RawButton := bench.Operator.JoyBtnRaw, Cfg := cfg, NeutralXMem := nx, NeutralYMem := ny);
home(DeadmanArmed := joy.DeadmanArmed, JoystickDeflected := NOT joy.AtNeutralXY, JoystickPull := joy.AxisCmdY.DirectionPositive, JoystickPush := joy.AxisCmdY.DirectionNegative, BtnValidation := bench.Operator.JoyBtnRaw);
IF bench.Operator.JoyBtnRaw AND NOT previousButton THEN buttonEdges := buttonEdges + 1; END_IF; previousButton := bench.Operator.JoyBtnRaw;
ADVANCE_TIME(10000000);
bench(RawPosM1 := raw1, RawPosM2 := raw2);
joy(RawX := bench.Operator.JoyXRaw_ANA1, RawY := bench.Operator.JoyYRaw_ANA2, RawButton := bench.Operator.JoyBtnRaw, Cfg := cfg, NeutralXMem := nx, NeutralYMem := ny);
home(DeadmanArmed := joy.DeadmanArmed, JoystickDeflected := NOT joy.AtNeutralXY, JoystickPull := joy.AxisCmdY.DirectionPositive, JoystickPush := joy.AxisCmdY.DirectionNegative, BtnValidation := bench.Operator.JoyBtnRaw);
IF bench.Operator.JoyBtnRaw AND NOT previousButton THEN buttonEdges := buttonEdges + 1; END_IF; previousButton := bench.Operator.JoyBtnRaw;
ADVANCE_TIME(10000000);
bench(RawPosM1 := raw1, RawPosM2 := raw2);
joy(RawX := bench.Operator.JoyXRaw_ANA1, RawY := bench.Operator.JoyYRaw_ANA2, RawButton := bench.Operator.JoyBtnRaw, Cfg := cfg, NeutralXMem := nx, NeutralYMem := ny);
home(DeadmanArmed := joy.DeadmanArmed, JoystickDeflected := NOT joy.AtNeutralXY, JoystickPull := joy.AxisCmdY.DirectionPositive, JoystickPush := joy.AxisCmdY.DirectionNegative, BtnValidation := bench.Operator.JoyBtnRaw);
IF bench.Operator.JoyBtnRaw AND NOT previousButton THEN buttonEdges := buttonEdges + 1; END_IF; previousButton := bench.Operator.JoyBtnRaw;
ADVANCE_TIME(10000000);
bench(RawPosM1 := raw1, RawPosM2 := raw2);
joy(RawX := bench.Operator.JoyXRaw_ANA1, RawY := bench.Operator.JoyYRaw_ANA2, RawButton := bench.Operator.JoyBtnRaw, Cfg := cfg, NeutralXMem := nx, NeutralYMem := ny);
home(DeadmanArmed := joy.DeadmanArmed, JoystickDeflected := NOT joy.AtNeutralXY, JoystickPull := joy.AxisCmdY.DirectionPositive, JoystickPush := joy.AxisCmdY.DirectionNegative, BtnValidation := bench.Operator.JoyBtnRaw);
IF bench.Operator.JoyBtnRaw AND NOT previousButton THEN buttonEdges := buttonEdges + 1; END_IF; previousButton := bench.Operator.JoyBtnRaw;
ADVANCE_TIME(10000000);
bench(RawPosM1 := raw1, RawPosM2 := raw2);
joy(RawX := bench.Operator.JoyXRaw_ANA1, RawY := bench.Operator.JoyYRaw_ANA2, RawButton := bench.Operator.JoyBtnRaw, Cfg := cfg, NeutralXMem := nx, NeutralYMem := ny);
home(DeadmanArmed := joy.DeadmanArmed, JoystickDeflected := NOT joy.AtNeutralXY, JoystickPull := joy.AxisCmdY.DirectionPositive, JoystickPush := joy.AxisCmdY.DirectionNegative, BtnValidation := bench.Operator.JoyBtnRaw);
IF bench.Operator.JoyBtnRaw AND NOT previousButton THEN buttonEdges := buttonEdges + 1; END_IF; previousButton := bench.Operator.JoyBtnRaw;
ADVANCE_TIME(10000000);
bench(RawPosM1 := raw1, RawPosM2 := raw2);
joy(RawX := bench.Operator.JoyXRaw_ANA1, RawY := bench.Operator.JoyYRaw_ANA2, RawButton := bench.Operator.JoyBtnRaw, Cfg := cfg, NeutralXMem := nx, NeutralYMem := ny);
home(DeadmanArmed := joy.DeadmanArmed, JoystickDeflected := NOT joy.AtNeutralXY, JoystickPull := joy.AxisCmdY.DirectionPositive, JoystickPush := joy.AxisCmdY.DirectionNegative, BtnValidation := bench.Operator.JoyBtnRaw);
IF bench.Operator.JoyBtnRaw AND NOT previousButton THEN buttonEdges := buttonEdges + 1; END_IF; previousButton := bench.Operator.JoyBtnRaw;
ADVANCE_TIME(10000000);
bench(RawPosM1 := raw1, RawPosM2 := raw2);
joy(RawX := bench.Operator.JoyXRaw_ANA1, RawY := bench.Operator.JoyYRaw_ANA2, RawButton := bench.Operator.JoyBtnRaw, Cfg := cfg, NeutralXMem := nx, NeutralYMem := ny);
home(DeadmanArmed := joy.DeadmanArmed, JoystickDeflected := NOT joy.AtNeutralXY, JoystickPull := joy.AxisCmdY.DirectionPositive, JoystickPush := joy.AxisCmdY.DirectionNegative, BtnValidation := bench.Operator.JoyBtnRaw);
IF bench.Operator.JoyBtnRaw AND NOT previousButton THEN buttonEdges := buttonEdges + 1; END_IF; previousButton := bench.Operator.JoyBtnRaw;
ADVANCE_TIME(10000000);
bench(RawPosM1 := raw1, RawPosM2 := raw2);
joy(RawX := bench.Operator.JoyXRaw_ANA1, RawY := bench.Operator.JoyYRaw_ANA2, RawButton := bench.Operator.JoyBtnRaw, Cfg := cfg, NeutralXMem := nx, NeutralYMem := ny);
home(DeadmanArmed := joy.DeadmanArmed, JoystickDeflected := NOT joy.AtNeutralXY, JoystickPull := joy.AxisCmdY.DirectionPositive, JoystickPush := joy.AxisCmdY.DirectionNegative, BtnValidation := bench.Operator.JoyBtnRaw);
IF bench.Operator.JoyBtnRaw AND NOT previousButton THEN buttonEdges := buttonEdges + 1; END_IF; previousButton := bench.Operator.JoyBtnRaw;
ADVANCE_TIME(10000000);
bench(RawPosM1 := raw1, RawPosM2 := raw2);
joy(RawX := bench.Operator.JoyXRaw_ANA1, RawY := bench.Operator.JoyYRaw_ANA2, RawButton := bench.Operator.JoyBtnRaw, Cfg := cfg, NeutralXMem := nx, NeutralYMem := ny);
home(DeadmanArmed := joy.DeadmanArmed, JoystickDeflected := NOT joy.AtNeutralXY, JoystickPull := joy.AxisCmdY.DirectionPositive, JoystickPush := joy.AxisCmdY.DirectionNegative, BtnValidation := bench.Operator.JoyBtnRaw);
IF bench.Operator.JoyBtnRaw AND NOT previousButton THEN buttonEdges := buttonEdges + 1; END_IF; previousButton := bench.Operator.JoyBtnRaw;
ADVANCE_TIME(10000000);
bench(RawPosM1 := raw1, RawPosM2 := raw2);
joy(RawX := bench.Operator.JoyXRaw_ANA1, RawY := bench.Operator.JoyYRaw_ANA2, RawButton := bench.Operator.JoyBtnRaw, Cfg := cfg, NeutralXMem := nx, NeutralYMem := ny);
home(DeadmanArmed := joy.DeadmanArmed, JoystickDeflected := NOT joy.AtNeutralXY, JoystickPull := joy.AxisCmdY.DirectionPositive, JoystickPush := joy.AxisCmdY.DirectionNegative, BtnValidation := bench.Operator.JoyBtnRaw);
IF bench.Operator.JoyBtnRaw AND NOT previousButton THEN buttonEdges := buttonEdges + 1; END_IF; previousButton := bench.Operator.JoyBtnRaw;
ADVANCE_TIME(10000000);
bench(RawPosM1 := raw1, RawPosM2 := raw2);
joy(RawX := bench.Operator.JoyXRaw_ANA1, RawY := bench.Operator.JoyYRaw_ANA2, RawButton := bench.Operator.JoyBtnRaw, Cfg := cfg, NeutralXMem := nx, NeutralYMem := ny);
home(DeadmanArmed := joy.DeadmanArmed, JoystickDeflected := NOT joy.AtNeutralXY, JoystickPull := joy.AxisCmdY.DirectionPositive, JoystickPush := joy.AxisCmdY.DirectionNegative, BtnValidation := bench.Operator.JoyBtnRaw);
IF bench.Operator.JoyBtnRaw AND NOT previousButton THEN buttonEdges := buttonEdges + 1; END_IF; previousButton := bench.Operator.JoyBtnRaw;
ADVANCE_TIME(10000000);
bench(RawPosM1 := raw1, RawPosM2 := raw2);
joy(RawX := bench.Operator.JoyXRaw_ANA1, RawY := bench.Operator.JoyYRaw_ANA2, RawButton := bench.Operator.JoyBtnRaw, Cfg := cfg, NeutralXMem := nx, NeutralYMem := ny);
home(DeadmanArmed := joy.DeadmanArmed, JoystickDeflected := NOT joy.AtNeutralXY, JoystickPull := joy.AxisCmdY.DirectionPositive, JoystickPush := joy.AxisCmdY.DirectionNegative, BtnValidation := bench.Operator.JoyBtnRaw);
IF bench.Operator.JoyBtnRaw AND NOT previousButton THEN buttonEdges := buttonEdges + 1; END_IF; previousButton := bench.Operator.JoyBtnRaw;
ADVANCE_TIME(10000000);
bench(RawPosM1 := raw1, RawPosM2 := raw2);
joy(RawX := bench.Operator.JoyXRaw_ANA1, RawY := bench.Operator.JoyYRaw_ANA2, RawButton := bench.Operator.JoyBtnRaw, Cfg := cfg, NeutralXMem := nx, NeutralYMem := ny);
home(DeadmanArmed := joy.DeadmanArmed, JoystickDeflected := NOT joy.AtNeutralXY, JoystickPull := joy.AxisCmdY.DirectionPositive, JoystickPush := joy.AxisCmdY.DirectionNegative, BtnValidation := bench.Operator.JoyBtnRaw);
IF bench.Operator.JoyBtnRaw AND NOT previousButton THEN buttonEdges := buttonEdges + 1; END_IF; previousButton := bench.Operator.JoyBtnRaw;
ADVANCE_TIME(10000000);
bench(RawPosM1 := raw1, RawPosM2 := raw2);
joy(RawX := bench.Operator.JoyXRaw_ANA1, RawY := bench.Operator.JoyYRaw_ANA2, RawButton := bench.Operator.JoyBtnRaw, Cfg := cfg, NeutralXMem := nx, NeutralYMem := ny);
home(DeadmanArmed := joy.DeadmanArmed, JoystickDeflected := NOT joy.AtNeutralXY, JoystickPull := joy.AxisCmdY.DirectionPositive, JoystickPush := joy.AxisCmdY.DirectionNegative, BtnValidation := bench.Operator.JoyBtnRaw);
IF bench.Operator.JoyBtnRaw AND NOT previousButton THEN buttonEdges := buttonEdges + 1; END_IF; previousButton := bench.Operator.JoyBtnRaw;
ADVANCE_TIME(10000000);
bench(RawPosM1 := raw1, RawPosM2 := raw2);
joy(RawX := bench.Operator.JoyXRaw_ANA1, RawY := bench.Operator.JoyYRaw_ANA2, RawButton := bench.Operator.JoyBtnRaw, Cfg := cfg, NeutralXMem := nx, NeutralYMem := ny);
home(DeadmanArmed := joy.DeadmanArmed, JoystickDeflected := NOT joy.AtNeutralXY, JoystickPull := joy.AxisCmdY.DirectionPositive, JoystickPush := joy.AxisCmdY.DirectionNegative, BtnValidation := bench.Operator.JoyBtnRaw);
IF bench.Operator.JoyBtnRaw AND NOT previousButton THEN buttonEdges := buttonEdges + 1; END_IF; previousButton := bench.Operator.JoyBtnRaw;
ADVANCE_TIME(10000000);
bench(RawPosM1 := raw1, RawPosM2 := raw2);
joy(RawX := bench.Operator.JoyXRaw_ANA1, RawY := bench.Operator.JoyYRaw_ANA2, RawButton := bench.Operator.JoyBtnRaw, Cfg := cfg, NeutralXMem := nx, NeutralYMem := ny);
home(DeadmanArmed := joy.DeadmanArmed, JoystickDeflected := NOT joy.AtNeutralXY, JoystickPull := joy.AxisCmdY.DirectionPositive, JoystickPush := joy.AxisCmdY.DirectionNegative, BtnValidation := bench.Operator.JoyBtnRaw);
IF bench.Operator.JoyBtnRaw AND NOT previousButton THEN buttonEdges := buttonEdges + 1; END_IF; previousButton := bench.Operator.JoyBtnRaw;
ADVANCE_TIME(10000000);
bench(RawPosM1 := raw1, RawPosM2 := raw2);
joy(RawX := bench.Operator.JoyXRaw_ANA1, RawY := bench.Operator.JoyYRaw_ANA2, RawButton := bench.Operator.JoyBtnRaw, Cfg := cfg, NeutralXMem := nx, NeutralYMem := ny);
home(DeadmanArmed := joy.DeadmanArmed, JoystickDeflected := NOT joy.AtNeutralXY, JoystickPull := joy.AxisCmdY.DirectionPositive, JoystickPush := joy.AxisCmdY.DirectionNegative, BtnValidation := bench.Operator.JoyBtnRaw);
IF bench.Operator.JoyBtnRaw AND NOT previousButton THEN buttonEdges := buttonEdges + 1; END_IF; previousButton := bench.Operator.JoyBtnRaw;
ADVANCE_TIME(10000000);
bench(RawPosM1 := raw1, RawPosM2 := raw2);
joy(RawX := bench.Operator.JoyXRaw_ANA1, RawY := bench.Operator.JoyYRaw_ANA2, RawButton := bench.Operator.JoyBtnRaw, Cfg := cfg, NeutralXMem := nx, NeutralYMem := ny);
home(DeadmanArmed := joy.DeadmanArmed, JoystickDeflected := NOT joy.AtNeutralXY, JoystickPull := joy.AxisCmdY.DirectionPositive, JoystickPush := joy.AxisCmdY.DirectionNegative, BtnValidation := bench.Operator.JoyBtnRaw);
IF bench.Operator.JoyBtnRaw AND NOT previousButton THEN buttonEdges := buttonEdges + 1; END_IF; previousButton := bench.Operator.JoyBtnRaw;
ADVANCE_TIME(10000000);
bench(RawPosM1 := raw1, RawPosM2 := raw2);
joy(RawX := bench.Operator.JoyXRaw_ANA1, RawY := bench.Operator.JoyYRaw_ANA2, RawButton := bench.Operator.JoyBtnRaw, Cfg := cfg, NeutralXMem := nx, NeutralYMem := ny);
home(DeadmanArmed := joy.DeadmanArmed, JoystickDeflected := NOT joy.AtNeutralXY, JoystickPull := joy.AxisCmdY.DirectionPositive, JoystickPush := joy.AxisCmdY.DirectionNegative, BtnValidation := bench.Operator.JoyBtnRaw);
IF bench.Operator.JoyBtnRaw AND NOT previousButton THEN buttonEdges := buttonEdges + 1; END_IF; previousButton := bench.Operator.JoyBtnRaw;
ADVANCE_TIME(10000000);
bench(RawPosM1 := raw1, RawPosM2 := raw2);
joy(RawX := bench.Operator.JoyXRaw_ANA1, RawY := bench.Operator.JoyYRaw_ANA2, RawButton := bench.Operator.JoyBtnRaw, Cfg := cfg, NeutralXMem := nx, NeutralYMem := ny);
home(DeadmanArmed := joy.DeadmanArmed, JoystickDeflected := NOT joy.AtNeutralXY, JoystickPull := joy.AxisCmdY.DirectionPositive, JoystickPush := joy.AxisCmdY.DirectionNegative, BtnValidation := bench.Operator.JoyBtnRaw);
IF bench.Operator.JoyBtnRaw AND NOT previousButton THEN buttonEdges := buttonEdges + 1; END_IF; previousButton := bench.Operator.JoyBtnRaw;
ADVANCE_TIME(10000000);
bench(RawPosM1 := raw1, RawPosM2 := raw2);
joy(RawX := bench.Operator.JoyXRaw_ANA1, RawY := bench.Operator.JoyYRaw_ANA2, RawButton := bench.Operator.JoyBtnRaw, Cfg := cfg, NeutralXMem := nx, NeutralYMem := ny);
home(DeadmanArmed := joy.DeadmanArmed, JoystickDeflected := NOT joy.AtNeutralXY, JoystickPull := joy.AxisCmdY.DirectionPositive, JoystickPush := joy.AxisCmdY.DirectionNegative, BtnValidation := bench.Operator.JoyBtnRaw);
IF bench.Operator.JoyBtnRaw AND NOT previousButton THEN buttonEdges := buttonEdges + 1; END_IF; previousButton := bench.Operator.JoyBtnRaw;
ADVANCE_TIME(10000000);
bench(RawPosM1 := raw1, RawPosM2 := raw2);
joy(RawX := bench.Operator.JoyXRaw_ANA1, RawY := bench.Operator.JoyYRaw_ANA2, RawButton := bench.Operator.JoyBtnRaw, Cfg := cfg, NeutralXMem := nx, NeutralYMem := ny);
home(DeadmanArmed := joy.DeadmanArmed, JoystickDeflected := NOT joy.AtNeutralXY, JoystickPull := joy.AxisCmdY.DirectionPositive, JoystickPush := joy.AxisCmdY.DirectionNegative, BtnValidation := bench.Operator.JoyBtnRaw);
IF bench.Operator.JoyBtnRaw AND NOT previousButton THEN buttonEdges := buttonEdges + 1; END_IF; previousButton := bench.Operator.JoyBtnRaw;
ADVANCE_TIME(10000000);
bench(RawPosM1 := raw1, RawPosM2 := raw2);
joy(RawX := bench.Operator.JoyXRaw_ANA1, RawY := bench.Operator.JoyYRaw_ANA2, RawButton := bench.Operator.JoyBtnRaw, Cfg := cfg, NeutralXMem := nx, NeutralYMem := ny);
home(DeadmanArmed := joy.DeadmanArmed, JoystickDeflected := NOT joy.AtNeutralXY, JoystickPull := joy.AxisCmdY.DirectionPositive, JoystickPush := joy.AxisCmdY.DirectionNegative, BtnValidation := bench.Operator.JoyBtnRaw);
IF bench.Operator.JoyBtnRaw AND NOT previousButton THEN buttonEdges := buttonEdges + 1; END_IF; previousButton := bench.Operator.JoyBtnRaw;
ADVANCE_TIME(10000000);
bench(RawPosM1 := raw1, RawPosM2 := raw2);
joy(RawX := bench.Operator.JoyXRaw_ANA1, RawY := bench.Operator.JoyYRaw_ANA2, RawButton := bench.Operator.JoyBtnRaw, Cfg := cfg, NeutralXMem := nx, NeutralYMem := ny);
home(DeadmanArmed := joy.DeadmanArmed, JoystickDeflected := NOT joy.AtNeutralXY, JoystickPull := joy.AxisCmdY.DirectionPositive, JoystickPush := joy.AxisCmdY.DirectionNegative, BtnValidation := bench.Operator.JoyBtnRaw);
IF bench.Operator.JoyBtnRaw AND NOT previousButton THEN buttonEdges := buttonEdges + 1; END_IF; previousButton := bench.Operator.JoyBtnRaw;
ADVANCE_TIME(10000000);
bench(RawPosM1 := raw1, RawPosM2 := raw2);
joy(RawX := bench.Operator.JoyXRaw_ANA1, RawY := bench.Operator.JoyYRaw_ANA2, RawButton := bench.Operator.JoyBtnRaw, Cfg := cfg, NeutralXMem := nx, NeutralYMem := ny);
home(DeadmanArmed := joy.DeadmanArmed, JoystickDeflected := NOT joy.AtNeutralXY, JoystickPull := joy.AxisCmdY.DirectionPositive, JoystickPush := joy.AxisCmdY.DirectionNegative, BtnValidation := bench.Operator.JoyBtnRaw);
IF bench.Operator.JoyBtnRaw AND NOT previousButton THEN buttonEdges := buttonEdges + 1; END_IF; previousButton := bench.Operator.JoyBtnRaw;
ADVANCE_TIME(10000000);
bench(RawPosM1 := raw1, RawPosM2 := raw2);
joy(RawX := bench.Operator.JoyXRaw_ANA1, RawY := bench.Operator.JoyYRaw_ANA2, RawButton := bench.Operator.JoyBtnRaw, Cfg := cfg, NeutralXMem := nx, NeutralYMem := ny);
home(DeadmanArmed := joy.DeadmanArmed, JoystickDeflected := NOT joy.AtNeutralXY, JoystickPull := joy.AxisCmdY.DirectionPositive, JoystickPush := joy.AxisCmdY.DirectionNegative, BtnValidation := bench.Operator.JoyBtnRaw);
IF bench.Operator.JoyBtnRaw AND NOT previousButton THEN buttonEdges := buttonEdges + 1; END_IF; previousButton := bench.Operator.JoyBtnRaw;
ADVANCE_TIME(10000000);
bench(RawPosM1 := raw1, RawPosM2 := raw2);
joy(RawX := bench.Operator.JoyXRaw_ANA1, RawY := bench.Operator.JoyYRaw_ANA2, RawButton := bench.Operator.JoyBtnRaw, Cfg := cfg, NeutralXMem := nx, NeutralYMem := ny);
home(DeadmanArmed := joy.DeadmanArmed, JoystickDeflected := NOT joy.AtNeutralXY, JoystickPull := joy.AxisCmdY.DirectionPositive, JoystickPush := joy.AxisCmdY.DirectionNegative, BtnValidation := bench.Operator.JoyBtnRaw);
IF bench.Operator.JoyBtnRaw AND NOT previousButton THEN buttonEdges := buttonEdges + 1; END_IF; previousButton := bench.Operator.JoyBtnRaw;
ADVANCE_TIME(10000000);
bench(RawPosM1 := raw1, RawPosM2 := raw2);
joy(RawX := bench.Operator.JoyXRaw_ANA1, RawY := bench.Operator.JoyYRaw_ANA2, RawButton := bench.Operator.JoyBtnRaw, Cfg := cfg, NeutralXMem := nx, NeutralYMem := ny);
home(DeadmanArmed := joy.DeadmanArmed, JoystickDeflected := NOT joy.AtNeutralXY, JoystickPull := joy.AxisCmdY.DirectionPositive, JoystickPush := joy.AxisCmdY.DirectionNegative, BtnValidation := bench.Operator.JoyBtnRaw);
IF bench.Operator.JoyBtnRaw AND NOT previousButton THEN buttonEdges := buttonEdges + 1; END_IF; previousButton := bench.Operator.JoyBtnRaw;
ADVANCE_TIME(10000000);
bench(RawPosM1 := raw1, RawPosM2 := raw2);
joy(RawX := bench.Operator.JoyXRaw_ANA1, RawY := bench.Operator.JoyYRaw_ANA2, RawButton := bench.Operator.JoyBtnRaw, Cfg := cfg, NeutralXMem := nx, NeutralYMem := ny);
home(DeadmanArmed := joy.DeadmanArmed, JoystickDeflected := NOT joy.AtNeutralXY, JoystickPull := joy.AxisCmdY.DirectionPositive, JoystickPush := joy.AxisCmdY.DirectionNegative, BtnValidation := bench.Operator.JoyBtnRaw);
IF bench.Operator.JoyBtnRaw AND NOT previousButton THEN buttonEdges := buttonEdges + 1; END_IF; previousButton := bench.Operator.JoyBtnRaw;
ADVANCE_TIME(10000000);
bench(RawPosM1 := raw1, RawPosM2 := raw2);
joy(RawX := bench.Operator.JoyXRaw_ANA1, RawY := bench.Operator.JoyYRaw_ANA2, RawButton := bench.Operator.JoyBtnRaw, Cfg := cfg, NeutralXMem := nx, NeutralYMem := ny);
home(DeadmanArmed := joy.DeadmanArmed, JoystickDeflected := NOT joy.AtNeutralXY, JoystickPull := joy.AxisCmdY.DirectionPositive, JoystickPush := joy.AxisCmdY.DirectionNegative, BtnValidation := bench.Operator.JoyBtnRaw);
IF bench.Operator.JoyBtnRaw AND NOT previousButton THEN buttonEdges := buttonEdges + 1; END_IF; previousButton := bench.Operator.JoyBtnRaw;
ADVANCE_TIME(10000000);
bench(RawPosM1 := raw1, RawPosM2 := raw2);
joy(RawX := bench.Operator.JoyXRaw_ANA1, RawY := bench.Operator.JoyYRaw_ANA2, RawButton := bench.Operator.JoyBtnRaw, Cfg := cfg, NeutralXMem := nx, NeutralYMem := ny);
home(DeadmanArmed := joy.DeadmanArmed, JoystickDeflected := NOT joy.AtNeutralXY, JoystickPull := joy.AxisCmdY.DirectionPositive, JoystickPush := joy.AxisCmdY.DirectionNegative, BtnValidation := bench.Operator.JoyBtnRaw);
IF bench.Operator.JoyBtnRaw AND NOT previousButton THEN buttonEdges := buttonEdges + 1; END_IF; previousButton := bench.Operator.JoyBtnRaw;
ADVANCE_TIME(10000000);
bench(RawPosM1 := raw1, RawPosM2 := raw2);
joy(RawX := bench.Operator.JoyXRaw_ANA1, RawY := bench.Operator.JoyYRaw_ANA2, RawButton := bench.Operator.JoyBtnRaw, Cfg := cfg, NeutralXMem := nx, NeutralYMem := ny);
home(DeadmanArmed := joy.DeadmanArmed, JoystickDeflected := NOT joy.AtNeutralXY, JoystickPull := joy.AxisCmdY.DirectionPositive, JoystickPush := joy.AxisCmdY.DirectionNegative, BtnValidation := bench.Operator.JoyBtnRaw);
IF bench.Operator.JoyBtnRaw AND NOT previousButton THEN buttonEdges := buttonEdges + 1; END_IF; previousButton := bench.Operator.JoyBtnRaw;
ASSERT_TRUE(joy.AxisCmdX.DirectionNegative, 'Second geste rapproche accepte par logique reelle'); ASSERT_EQ(buttonEdges, 2, 'Un front par geste');
bench.SimJoystickLeft_Rev_TREMIE_Active := FALSE;
ADVANCE_TIME(10000000);
bench(RawPosM1 := raw1, RawPosM2 := raw2);
joy(RawX := bench.Operator.JoyXRaw_ANA1, RawY := bench.Operator.JoyYRaw_ANA2, RawButton := bench.Operator.JoyBtnRaw, Cfg := cfg, NeutralXMem := nx, NeutralYMem := ny);
home(DeadmanArmed := joy.DeadmanArmed, JoystickDeflected := NOT joy.AtNeutralXY, JoystickPull := joy.AxisCmdY.DirectionPositive, JoystickPush := joy.AxisCmdY.DirectionNegative, BtnValidation := bench.Operator.JoyBtnRaw);
IF bench.Operator.JoyBtnRaw AND NOT previousButton THEN buttonEdges := buttonEdges + 1; END_IF; previousButton := bench.Operator.JoyBtnRaw;
ADVANCE_TIME(10000000);
bench(RawPosM1 := raw1, RawPosM2 := raw2);
joy(RawX := bench.Operator.JoyXRaw_ANA1, RawY := bench.Operator.JoyYRaw_ANA2, RawButton := bench.Operator.JoyBtnRaw, Cfg := cfg, NeutralXMem := nx, NeutralYMem := ny);
home(DeadmanArmed := joy.DeadmanArmed, JoystickDeflected := NOT joy.AtNeutralXY, JoystickPull := joy.AxisCmdY.DirectionPositive, JoystickPush := joy.AxisCmdY.DirectionNegative, BtnValidation := bench.Operator.JoyBtnRaw);
IF bench.Operator.JoyBtnRaw AND NOT previousButton THEN buttonEdges := buttonEdges + 1; END_IF; previousButton := bench.Operator.JoyBtnRaw;
ADVANCE_TIME(10000000);
bench(RawPosM1 := raw1, RawPosM2 := raw2);
joy(RawX := bench.Operator.JoyXRaw_ANA1, RawY := bench.Operator.JoyYRaw_ANA2, RawButton := bench.Operator.JoyBtnRaw, Cfg := cfg, NeutralXMem := nx, NeutralYMem := ny);
home(DeadmanArmed := joy.DeadmanArmed, JoystickDeflected := NOT joy.AtNeutralXY, JoystickPull := joy.AxisCmdY.DirectionPositive, JoystickPush := joy.AxisCmdY.DirectionNegative, BtnValidation := bench.Operator.JoyBtnRaw);
IF bench.Operator.JoyBtnRaw AND NOT previousButton THEN buttonEdges := buttonEdges + 1; END_IF; previousButton := bench.Operator.JoyBtnRaw;
ADVANCE_TIME(10000000);
bench(RawPosM1 := raw1, RawPosM2 := raw2);
joy(RawX := bench.Operator.JoyXRaw_ANA1, RawY := bench.Operator.JoyYRaw_ANA2, RawButton := bench.Operator.JoyBtnRaw, Cfg := cfg, NeutralXMem := nx, NeutralYMem := ny);
home(DeadmanArmed := joy.DeadmanArmed, JoystickDeflected := NOT joy.AtNeutralXY, JoystickPull := joy.AxisCmdY.DirectionPositive, JoystickPush := joy.AxisCmdY.DirectionNegative, BtnValidation := bench.Operator.JoyBtnRaw);
IF bench.Operator.JoyBtnRaw AND NOT previousButton THEN buttonEdges := buttonEdges + 1; END_IF; previousButton := bench.Operator.JoyBtnRaw;
ADVANCE_TIME(10000000);
bench(RawPosM1 := raw1, RawPosM2 := raw2);
joy(RawX := bench.Operator.JoyXRaw_ANA1, RawY := bench.Operator.JoyYRaw_ANA2, RawButton := bench.Operator.JoyBtnRaw, Cfg := cfg, NeutralXMem := nx, NeutralYMem := ny);
home(DeadmanArmed := joy.DeadmanArmed, JoystickDeflected := NOT joy.AtNeutralXY, JoystickPull := joy.AxisCmdY.DirectionPositive, JoystickPush := joy.AxisCmdY.DirectionNegative, BtnValidation := bench.Operator.JoyBtnRaw);
IF bench.Operator.JoyBtnRaw AND NOT previousButton THEN buttonEdges := buttonEdges + 1; END_IF; previousButton := bench.Operator.JoyBtnRaw;
ADVANCE_TIME(10000000);
bench(RawPosM1 := raw1, RawPosM2 := raw2);
joy(RawX := bench.Operator.JoyXRaw_ANA1, RawY := bench.Operator.JoyYRaw_ANA2, RawButton := bench.Operator.JoyBtnRaw, Cfg := cfg, NeutralXMem := nx, NeutralYMem := ny);
home(DeadmanArmed := joy.DeadmanArmed, JoystickDeflected := NOT joy.AtNeutralXY, JoystickPull := joy.AxisCmdY.DirectionPositive, JoystickPush := joy.AxisCmdY.DirectionNegative, BtnValidation := bench.Operator.JoyBtnRaw);
IF bench.Operator.JoyBtnRaw AND NOT previousButton THEN buttonEdges := buttonEdges + 1; END_IF; previousButton := bench.Operator.JoyBtnRaw;
ADVANCE_TIME(10000000);
bench(RawPosM1 := raw1, RawPosM2 := raw2);
joy(RawX := bench.Operator.JoyXRaw_ANA1, RawY := bench.Operator.JoyYRaw_ANA2, RawButton := bench.Operator.JoyBtnRaw, Cfg := cfg, NeutralXMem := nx, NeutralYMem := ny);
home(DeadmanArmed := joy.DeadmanArmed, JoystickDeflected := NOT joy.AtNeutralXY, JoystickPull := joy.AxisCmdY.DirectionPositive, JoystickPush := joy.AxisCmdY.DirectionNegative, BtnValidation := bench.Operator.JoyBtnRaw);
IF bench.Operator.JoyBtnRaw AND NOT previousButton THEN buttonEdges := buttonEdges + 1; END_IF; previousButton := bench.Operator.JoyBtnRaw;
ADVANCE_TIME(10000000);
bench(RawPosM1 := raw1, RawPosM2 := raw2);
joy(RawX := bench.Operator.JoyXRaw_ANA1, RawY := bench.Operator.JoyYRaw_ANA2, RawButton := bench.Operator.JoyBtnRaw, Cfg := cfg, NeutralXMem := nx, NeutralYMem := ny);
home(DeadmanArmed := joy.DeadmanArmed, JoystickDeflected := NOT joy.AtNeutralXY, JoystickPull := joy.AxisCmdY.DirectionPositive, JoystickPush := joy.AxisCmdY.DirectionNegative, BtnValidation := bench.Operator.JoyBtnRaw);
IF bench.Operator.JoyBtnRaw AND NOT previousButton THEN buttonEdges := buttonEdges + 1; END_IF; previousButton := bench.Operator.JoyBtnRaw;
ADVANCE_TIME(10000000);
bench(RawPosM1 := raw1, RawPosM2 := raw2);
joy(RawX := bench.Operator.JoyXRaw_ANA1, RawY := bench.Operator.JoyYRaw_ANA2, RawButton := bench.Operator.JoyBtnRaw, Cfg := cfg, NeutralXMem := nx, NeutralYMem := ny);
home(DeadmanArmed := joy.DeadmanArmed, JoystickDeflected := NOT joy.AtNeutralXY, JoystickPull := joy.AxisCmdY.DirectionPositive, JoystickPush := joy.AxisCmdY.DirectionNegative, BtnValidation := bench.Operator.JoyBtnRaw);
IF bench.Operator.JoyBtnRaw AND NOT previousButton THEN buttonEdges := buttonEdges + 1; END_IF; previousButton := bench.Operator.JoyBtnRaw;
ADVANCE_TIME(10000000);
bench(RawPosM1 := raw1, RawPosM2 := raw2);
joy(RawX := bench.Operator.JoyXRaw_ANA1, RawY := bench.Operator.JoyYRaw_ANA2, RawButton := bench.Operator.JoyBtnRaw, Cfg := cfg, NeutralXMem := nx, NeutralYMem := ny);
home(DeadmanArmed := joy.DeadmanArmed, JoystickDeflected := NOT joy.AtNeutralXY, JoystickPull := joy.AxisCmdY.DirectionPositive, JoystickPush := joy.AxisCmdY.DirectionNegative, BtnValidation := bench.Operator.JoyBtnRaw);
IF bench.Operator.JoyBtnRaw AND NOT previousButton THEN buttonEdges := buttonEdges + 1; END_IF; previousButton := bench.Operator.JoyBtnRaw;
ADVANCE_TIME(10000000);
bench(RawPosM1 := raw1, RawPosM2 := raw2);
joy(RawX := bench.Operator.JoyXRaw_ANA1, RawY := bench.Operator.JoyYRaw_ANA2, RawButton := bench.Operator.JoyBtnRaw, Cfg := cfg, NeutralXMem := nx, NeutralYMem := ny);
home(DeadmanArmed := joy.DeadmanArmed, JoystickDeflected := NOT joy.AtNeutralXY, JoystickPull := joy.AxisCmdY.DirectionPositive, JoystickPush := joy.AxisCmdY.DirectionNegative, BtnValidation := bench.Operator.JoyBtnRaw);
IF bench.Operator.JoyBtnRaw AND NOT previousButton THEN buttonEdges := buttonEdges + 1; END_IF; previousButton := bench.Operator.JoyBtnRaw;
ADVANCE_TIME(10000000);
bench(RawPosM1 := raw1, RawPosM2 := raw2);
joy(RawX := bench.Operator.JoyXRaw_ANA1, RawY := bench.Operator.JoyYRaw_ANA2, RawButton := bench.Operator.JoyBtnRaw, Cfg := cfg, NeutralXMem := nx, NeutralYMem := ny);
home(DeadmanArmed := joy.DeadmanArmed, JoystickDeflected := NOT joy.AtNeutralXY, JoystickPull := joy.AxisCmdY.DirectionPositive, JoystickPush := joy.AxisCmdY.DirectionNegative, BtnValidation := bench.Operator.JoyBtnRaw);
IF bench.Operator.JoyBtnRaw AND NOT previousButton THEN buttonEdges := buttonEdges + 1; END_IF; previousButton := bench.Operator.JoyBtnRaw;
ADVANCE_TIME(10000000);
bench(RawPosM1 := raw1, RawPosM2 := raw2);
joy(RawX := bench.Operator.JoyXRaw_ANA1, RawY := bench.Operator.JoyYRaw_ANA2, RawButton := bench.Operator.JoyBtnRaw, Cfg := cfg, NeutralXMem := nx, NeutralYMem := ny);
home(DeadmanArmed := joy.DeadmanArmed, JoystickDeflected := NOT joy.AtNeutralXY, JoystickPull := joy.AxisCmdY.DirectionPositive, JoystickPush := joy.AxisCmdY.DirectionNegative, BtnValidation := bench.Operator.JoyBtnRaw);
IF bench.Operator.JoyBtnRaw AND NOT previousButton THEN buttonEdges := buttonEdges + 1; END_IF; previousButton := bench.Operator.JoyBtnRaw;
ADVANCE_TIME(10000000);
bench(RawPosM1 := raw1, RawPosM2 := raw2);
joy(RawX := bench.Operator.JoyXRaw_ANA1, RawY := bench.Operator.JoyYRaw_ANA2, RawButton := bench.Operator.JoyBtnRaw, Cfg := cfg, NeutralXMem := nx, NeutralYMem := ny);
home(DeadmanArmed := joy.DeadmanArmed, JoystickDeflected := NOT joy.AtNeutralXY, JoystickPull := joy.AxisCmdY.DirectionPositive, JoystickPush := joy.AxisCmdY.DirectionNegative, BtnValidation := bench.Operator.JoyBtnRaw);
IF bench.Operator.JoyBtnRaw AND NOT previousButton THEN buttonEdges := buttonEdges + 1; END_IF; previousButton := bench.Operator.JoyBtnRaw;
ADVANCE_TIME(10000000);
bench(RawPosM1 := raw1, RawPosM2 := raw2);
joy(RawX := bench.Operator.JoyXRaw_ANA1, RawY := bench.Operator.JoyYRaw_ANA2, RawButton := bench.Operator.JoyBtnRaw, Cfg := cfg, NeutralXMem := nx, NeutralYMem := ny);
home(DeadmanArmed := joy.DeadmanArmed, JoystickDeflected := NOT joy.AtNeutralXY, JoystickPull := joy.AxisCmdY.DirectionPositive, JoystickPush := joy.AxisCmdY.DirectionNegative, BtnValidation := bench.Operator.JoyBtnRaw);
IF bench.Operator.JoyBtnRaw AND NOT previousButton THEN buttonEdges := buttonEdges + 1; END_IF; previousButton := bench.Operator.JoyBtnRaw;
ADVANCE_TIME(10000000);
bench(RawPosM1 := raw1, RawPosM2 := raw2);
joy(RawX := bench.Operator.JoyXRaw_ANA1, RawY := bench.Operator.JoyYRaw_ANA2, RawButton := bench.Operator.JoyBtnRaw, Cfg := cfg, NeutralXMem := nx, NeutralYMem := ny);
home(DeadmanArmed := joy.DeadmanArmed, JoystickDeflected := NOT joy.AtNeutralXY, JoystickPull := joy.AxisCmdY.DirectionPositive, JoystickPush := joy.AxisCmdY.DirectionNegative, BtnValidation := bench.Operator.JoyBtnRaw);
IF bench.Operator.JoyBtnRaw AND NOT previousButton THEN buttonEdges := buttonEdges + 1; END_IF; previousButton := bench.Operator.JoyBtnRaw;
ADVANCE_TIME(10000000);
bench(RawPosM1 := raw1, RawPosM2 := raw2);
joy(RawX := bench.Operator.JoyXRaw_ANA1, RawY := bench.Operator.JoyYRaw_ANA2, RawButton := bench.Operator.JoyBtnRaw, Cfg := cfg, NeutralXMem := nx, NeutralYMem := ny);
home(DeadmanArmed := joy.DeadmanArmed, JoystickDeflected := NOT joy.AtNeutralXY, JoystickPull := joy.AxisCmdY.DirectionPositive, JoystickPush := joy.AxisCmdY.DirectionNegative, BtnValidation := bench.Operator.JoyBtnRaw);
IF bench.Operator.JoyBtnRaw AND NOT previousButton THEN buttonEdges := buttonEdges + 1; END_IF; previousButton := bench.Operator.JoyBtnRaw;
ADVANCE_TIME(10000000);
bench(RawPosM1 := raw1, RawPosM2 := raw2);
joy(RawX := bench.Operator.JoyXRaw_ANA1, RawY := bench.Operator.JoyYRaw_ANA2, RawButton := bench.Operator.JoyBtnRaw, Cfg := cfg, NeutralXMem := nx, NeutralYMem := ny);
home(DeadmanArmed := joy.DeadmanArmed, JoystickDeflected := NOT joy.AtNeutralXY, JoystickPull := joy.AxisCmdY.DirectionPositive, JoystickPush := joy.AxisCmdY.DirectionNegative, BtnValidation := bench.Operator.JoyBtnRaw);
IF bench.Operator.JoyBtnRaw AND NOT previousButton THEN buttonEdges := buttonEdges + 1; END_IF; previousButton := bench.Operator.JoyBtnRaw;
ADVANCE_TIME(10000000);
bench(RawPosM1 := raw1, RawPosM2 := raw2);
joy(RawX := bench.Operator.JoyXRaw_ANA1, RawY := bench.Operator.JoyYRaw_ANA2, RawButton := bench.Operator.JoyBtnRaw, Cfg := cfg, NeutralXMem := nx, NeutralYMem := ny);
home(DeadmanArmed := joy.DeadmanArmed, JoystickDeflected := NOT joy.AtNeutralXY, JoystickPull := joy.AxisCmdY.DirectionPositive, JoystickPush := joy.AxisCmdY.DirectionNegative, BtnValidation := bench.Operator.JoyBtnRaw);
IF bench.Operator.JoyBtnRaw AND NOT previousButton THEN buttonEdges := buttonEdges + 1; END_IF; previousButton := bench.Operator.JoyBtnRaw;
ADVANCE_TIME(10000000);
bench(RawPosM1 := raw1, RawPosM2 := raw2);
joy(RawX := bench.Operator.JoyXRaw_ANA1, RawY := bench.Operator.JoyYRaw_ANA2, RawButton := bench.Operator.JoyBtnRaw, Cfg := cfg, NeutralXMem := nx, NeutralYMem := ny);
home(DeadmanArmed := joy.DeadmanArmed, JoystickDeflected := NOT joy.AtNeutralXY, JoystickPull := joy.AxisCmdY.DirectionPositive, JoystickPush := joy.AxisCmdY.DirectionNegative, BtnValidation := bench.Operator.JoyBtnRaw);
IF bench.Operator.JoyBtnRaw AND NOT previousButton THEN buttonEdges := buttonEdges + 1; END_IF; previousButton := bench.Operator.JoyBtnRaw;
ADVANCE_TIME(10000000);
bench(RawPosM1 := raw1, RawPosM2 := raw2);
joy(RawX := bench.Operator.JoyXRaw_ANA1, RawY := bench.Operator.JoyYRaw_ANA2, RawButton := bench.Operator.JoyBtnRaw, Cfg := cfg, NeutralXMem := nx, NeutralYMem := ny);
home(DeadmanArmed := joy.DeadmanArmed, JoystickDeflected := NOT joy.AtNeutralXY, JoystickPull := joy.AxisCmdY.DirectionPositive, JoystickPush := joy.AxisCmdY.DirectionNegative, BtnValidation := bench.Operator.JoyBtnRaw);
IF bench.Operator.JoyBtnRaw AND NOT previousButton THEN buttonEdges := buttonEdges + 1; END_IF; previousButton := bench.Operator.JoyBtnRaw;
ADVANCE_TIME(10000000);
bench(RawPosM1 := raw1, RawPosM2 := raw2);
joy(RawX := bench.Operator.JoyXRaw_ANA1, RawY := bench.Operator.JoyYRaw_ANA2, RawButton := bench.Operator.JoyBtnRaw, Cfg := cfg, NeutralXMem := nx, NeutralYMem := ny);
home(DeadmanArmed := joy.DeadmanArmed, JoystickDeflected := NOT joy.AtNeutralXY, JoystickPull := joy.AxisCmdY.DirectionPositive, JoystickPush := joy.AxisCmdY.DirectionNegative, BtnValidation := bench.Operator.JoyBtnRaw);
IF bench.Operator.JoyBtnRaw AND NOT previousButton THEN buttonEdges := buttonEdges + 1; END_IF; previousButton := bench.Operator.JoyBtnRaw;
ADVANCE_TIME(10000000);
bench(RawPosM1 := raw1, RawPosM2 := raw2);
joy(RawX := bench.Operator.JoyXRaw_ANA1, RawY := bench.Operator.JoyYRaw_ANA2, RawButton := bench.Operator.JoyBtnRaw, Cfg := cfg, NeutralXMem := nx, NeutralYMem := ny);
home(DeadmanArmed := joy.DeadmanArmed, JoystickDeflected := NOT joy.AtNeutralXY, JoystickPull := joy.AxisCmdY.DirectionPositive, JoystickPush := joy.AxisCmdY.DirectionNegative, BtnValidation := bench.Operator.JoyBtnRaw);
IF bench.Operator.JoyBtnRaw AND NOT previousButton THEN buttonEdges := buttonEdges + 1; END_IF; previousButton := bench.Operator.JoyBtnRaw;
ADVANCE_TIME(10000000);
bench(RawPosM1 := raw1, RawPosM2 := raw2);
joy(RawX := bench.Operator.JoyXRaw_ANA1, RawY := bench.Operator.JoyYRaw_ANA2, RawButton := bench.Operator.JoyBtnRaw, Cfg := cfg, NeutralXMem := nx, NeutralYMem := ny);
home(DeadmanArmed := joy.DeadmanArmed, JoystickDeflected := NOT joy.AtNeutralXY, JoystickPull := joy.AxisCmdY.DirectionPositive, JoystickPush := joy.AxisCmdY.DirectionNegative, BtnValidation := bench.Operator.JoyBtnRaw);
IF bench.Operator.JoyBtnRaw AND NOT previousButton THEN buttonEdges := buttonEdges + 1; END_IF; previousButton := bench.Operator.JoyBtnRaw;
ADVANCE_TIME(10000000);
bench(RawPosM1 := raw1, RawPosM2 := raw2);
joy(RawX := bench.Operator.JoyXRaw_ANA1, RawY := bench.Operator.JoyYRaw_ANA2, RawButton := bench.Operator.JoyBtnRaw, Cfg := cfg, NeutralXMem := nx, NeutralYMem := ny);
home(DeadmanArmed := joy.DeadmanArmed, JoystickDeflected := NOT joy.AtNeutralXY, JoystickPull := joy.AxisCmdY.DirectionPositive, JoystickPush := joy.AxisCmdY.DirectionNegative, BtnValidation := bench.Operator.JoyBtnRaw);
IF bench.Operator.JoyBtnRaw AND NOT previousButton THEN buttonEdges := buttonEdges + 1; END_IF; previousButton := bench.Operator.JoyBtnRaw;
ADVANCE_TIME(4000000000);
ADVANCE_TIME(10000000);
bench(RawPosM1 := raw1, RawPosM2 := raw2);
joy(RawX := bench.Operator.JoyXRaw_ANA1, RawY := bench.Operator.JoyYRaw_ANA2, RawButton := bench.Operator.JoyBtnRaw, Cfg := cfg, NeutralXMem := nx, NeutralYMem := ny);
home(DeadmanArmed := joy.DeadmanArmed, JoystickDeflected := NOT joy.AtNeutralXY, JoystickPull := joy.AxisCmdY.DirectionPositive, JoystickPush := joy.AxisCmdY.DirectionNegative, BtnValidation := bench.Operator.JoyBtnRaw);
IF bench.Operator.JoyBtnRaw AND NOT previousButton THEN buttonEdges := buttonEdges + 1; END_IF; previousButton := bench.Operator.JoyBtnRaw;
ADVANCE_TIME(110000000);
ADVANCE_TIME(10000000);
bench(RawPosM1 := raw1, RawPosM2 := raw2);
joy(RawX := bench.Operator.JoyXRaw_ANA1, RawY := bench.Operator.JoyYRaw_ANA2, RawButton := bench.Operator.JoyBtnRaw, Cfg := cfg, NeutralXMem := nx, NeutralYMem := ny);
home(DeadmanArmed := joy.DeadmanArmed, JoystickDeflected := NOT joy.AtNeutralXY, JoystickPull := joy.AxisCmdY.DirectionPositive, JoystickPush := joy.AxisCmdY.DirectionNegative, BtnValidation := bench.Operator.JoyBtnRaw);
IF bench.Operator.JoyBtnRaw AND NOT previousButton THEN buttonEdges := buttonEdges + 1; END_IF; previousButton := bench.Operator.JoyBtnRaw;
ASSERT_FALSE(joy.DeadmanArmed, 'Desarmement reel apres grace et neutre');
END_TEST
